                    movel(spat_flatM_pick_p, a=0.2, v=0.1)
                    # begin: URCap Program Node
                    #   Source: Robotiq_Grippers, 3.17.0.105337, Robotiq Inc.
                    #   Type: Gripper
                    $ 4563 "Gripper Open (1)" "noBreak"
                    if not(gripper_connected[0]):
                      popup("Gripper 1 must be connected to run this program.", "No connection", False, True, True)
                    end
                    if not(rq_is_gripper_activated("1")):
                      popup("Gripper 1 is not activated. Go to Installation tab > Gripper to activate it and run the program again.", "Not activated", False, True, True)
                    end
                    rq_set_pos_spd_for(0, 0, 77, "1")
                    rq_wait_pos_spe_for_request(0, 0, 77, "1")
                    rq_go_to("1")
                    rq_wait("1")
                    # end: URCap Program Node
                    $ 4564 "spat_flatS_pick" "noBreak"
                    movel(spat_flatS_pick_p, a=1.2, v=0.25)
                    # begin: URCap Program Node
                    #   Source: Robotiq_Grippers, 3.17.0.105337, Robotiq Inc.
                    #   Type: Gripper
                    $ 4565 "Gripper Close (1)" "noBreak"
                    if not(gripper_connected[0]):
                      popup("Gripper 1 must be connected to run this program.", "No connection", False, True, True)
                    end
                    if not(rq_is_gripper_activated("1")):
                      popup("Gripper 1 is not activated. Go to Installation tab > Gripper to activate it and run the program again.", "Not activated", False, True, True)
                    end
                    rq_set_pos_spd_for(255, 0, 77, "1")
                    rq_wait_pos_spe_for_request(255, 0, 77, "1")
                    rq_go_to("1")
                    rq_wait("1")
                    # end: URCap Program Node
                    $ 4566 "spat_flatS_up" "noBreak"
                    movel(spat_flatS_up_p, a=1.2, v=0.25)
                    $ 4567 "Spatula_otw" "noBreak"
                    movel(Spatula_otw_p, a=1.2, v=0.25)
                    $ 4568 "switch_spat_F_S≔ False " "noBreak"
                    global switch_spat_F_S=  False
                    $ 4569 "correction_reset()" "noBreak"
                    correction_reset()
                  end
                end
              end
            end
            $ 4570 "tilt(level)" "noBreak"
            tilt(level)
            $ 4571 "Action_Info≔'Scooping'" "noBreak"
            global Action_Info="Scooping"
            $ 4572 "auto_tilt_and_scoop(W_now, target_weight, weight_value)" "noBreak"
            auto_tilt_and_scoop(W_now, target_weight, weight_value)
            $ 4573 "Action_Info≔'Dosing'" "noBreak"
            global Action_Info="Dosing"
          end
        end
        if (weight_value <= target_weight and delta_count<3):
          global thread_handler_4490=run Thread_while_4490()
          while (weight_value <= target_weight and delta_count<3):
            sync()
          end
          kill thread_handler_4490
        end
        # begin: URCap Program Node
        #   Source: SensoPart VISOR Robotic, 2.0.6, SensoPart Industriesensorik GmbH
        #   Type: Exit Pose
        $ 4574 "Exit Pose" "noBreak"
        movel(pose_trans(easyPickPose,p[0.0000,0.0000,-0.0000,0.0000,0.0000,0.0000]),a=0.5000,v=0.2500,t=0.000000,r=0.000000)
        # end: URCap Program Node
        easyPickObjTaken = True
      end
      # end: URCap Program Node
      # begin: URCap Program Node
      #   Source: SensoPart VISOR Robotic, 2.0.6, SensoPart Industriesensorik GmbH
      #   Type: No Object Detected
      $ 4575 "No Object Detected" "noBreak"
      if (visor_partsFound(easyPickVisorId) < 1):
        $ 4576 "Popup: No weigh scale detected" "noBreak"
        popup("No weigh scale detected", "Message", False, False, blocking=True)
        else:
      end
      # end: URCap Program Node
    end
    easyPickCount_4 = easyPickCount_4 + 1
    visor_easyPickUpdate(easyPickVisorId, "counter", easyPickCount_4)
    visor_easyPickSetIdent("bfde9f", easyPickVisorId)
    # end: URCap Program Node
  end
  visorFuncEasyPick_8737ac()
  # end: URCap Program Node
  $ 4577 "MoveL"
  $ 4578 "dispense_pos" "breakAfter"
  movel(dispense_pos, a=0.2, v=0.1)
  $ 4580 "Place spatula back to the rack"
  $ 4581 "If spatula ≟ 'spatula_L'"
  if (spatula  ==  "spatula_L"):
    $ 4582 "MoveJ"
    $ 4583 "Spatula_otw" "breakAfter"
    movej(get_inverse_kin(Spatula_otw_p, qnear=Spatula_otw_q), a=1.3962634015954636, v=1.0471975511965976)
    $ 4584 "MoveL"
    $ 4585 "spat_L_up" "breakAfter"
    movel(spat_L_up_p, a=1.2, v=0.25, r=0.05)
    $ 4586 "spat_L_side" "breakAfter"
    movel(spat_L_side_p, a=1.2, v=0.25, r=0.01)
    $ 4587 "spat_L_lift" "breakAfter"
    movel(spat_L_lift_p, a=1.2, v=0.25, r=0.01)
    $ 4588 "spat_L_pick" "breakAfter"
    movel(spat_L_pick_p, a=0.2, v=0.1)
    # begin: URCap Program Node
    #   Source: Robotiq_Grippers, 3.17.0.105337, Robotiq Inc.
    #   Type: Gripper
    $ 4589 "Gripper Open (1)"
    if not(gripper_connected[0]):
      popup("Gripper 1 must be connected to run this program.", "No connection", False, True, True)
    end
    if not(rq_is_gripper_activated("1")):
      popup("Gripper 1 is not activated. Go to Installation tab > Gripper to activate it and run the program again.", "Not activated", False, True, True)
    end
    rq_set_pos_spd_for(0, 128, 128, "1")
    rq_wait_pos_spe_for_request(0, 128, 128, "1")
    rq_go_to("1")
    rq_wait("1")
    # end: URCap Program Node
    $ 4590 "MoveJ"
    $ 4591 "pick_spat_L_abv" "breakAfter"
    movej(get_inverse_kin(pick_spat_L_abv_p, qnear=pick_spat_L_abv_q), a=1.3962634015954636, v=1.0471975511965976)
    $ 4592 "Spatula_otw" "breakAfter"
    movej(get_inverse_kin(Spatula_otw_p, qnear=Spatula_otw_q), a=1.3962634015954636, v=1.0471975511965976)
  else:
    $ 4593 "ElseIf spatula ≟'spatula_M'"
    if (spatula  == "spatula_M"):
      $ 4594 "MoveJ"
      $ 4595 "Spatula_otw" "breakAfter"
      movej(get_inverse_kin(Spatula_otw_p, qnear=Spatula_otw_q), a=1.3962634015954636, v=1.0471975511965976)
      $ 4596 "spat_M_up" "breakAfter"
      movej(get_inverse_kin(spat_M_up_p, qnear=spat_M_up_q), a=1.3962634015954636, v=1.0471975511965976, r=0.05)
      $ 4597 "MoveL"
      $ 4598 "spat_M_pick" "breakAfter"
      movel(spat_M_pick_p, a=0.2, v=0.1)
      # begin: URCap Program Node
      #   Source: Robotiq_Grippers, 3.17.0.105337, Robotiq Inc.
      #   Type: Gripper
      $ 4599 "Gripper Open (1)"
      if not(gripper_connected[0]):
        popup("Gripper 1 must be connected to run this program.", "No connection", False, True, True)
      end
      if not(rq_is_gripper_activated("1")):
        popup("Gripper 1 is not activated. Go to Installation tab > Gripper to activate it and run the program again.", "Not activated", False, True, True)
      end
      rq_set_pos_spd_for(0, 128, 128, "1")
      rq_wait_pos_spe_for_request(0, 128, 128, "1")
      rq_go_to("1")
      rq_wait("1")
      # end: URCap Program Node
      $ 4600 "spat_M_up" "breakAfter"
      movel(spat_M_up_p, a=1.2, v=0.25, r=0.05)
      $ 4601 "Spatula_otw" "breakAfter"
      movel(Spatula_otw_p, a=1.2, v=0.25)
      $ 4602 "switch_spat_M≔ False "
      global switch_spat_M=  False
    else:
      $ 4603 "ElseIf spatula≟'spatula_S'"
      if (spatula == "spatula_S"):
        $ 4604 "MoveJ"
        $ 4605 "Spatula_otw" "breakAfter"
        movej(get_inverse_kin(Spatula_otw_p, qnear=Spatula_otw_q), a=1.3962634015954636, v=1.0471975511965976)
        $ 4606 "spat_S_Up_7" "breakAfter"
        movej(get_inverse_kin(spat_S_Up_7_p, qnear=spat_S_Up_7_q), a=1.3962634015954636, v=1.0471975511965976, r=0.05)
        $ 4607 "MoveL"
        $ 4608 "spat_S_Pick_4" "breakAfter"
        movel(spat_S_Pick_4_p, a=0.2, v=0.1)
        # begin: URCap Program Node
        #   Source: Robotiq_Grippers, 3.17.0.105337, Robotiq Inc.
        #   Type: Gripper
        $ 4609 "Gripper Open (1)"
        if not(gripper_connected[0]):
          popup("Gripper 1 must be connected to run this program.", "No connection", False, True, True)
        end
        if not(rq_is_gripper_activated("1")):
          popup("Gripper 1 is not activated. Go to Installation tab > Gripper to activate it and run the program again.", "Not activated", False, True, True)
        end
        rq_set_pos_spd_for(0, 255, 51, "1")
        rq_wait_pos_spe_for_request(0, 255, 51, "1")
        rq_go_to("1")
        rq_wait("1")
        # end: URCap Program Node
        $ 4610 "spat_S_Up_8" "breakAfter"
        movel(spat_S_Up_8_p, a=1.2, v=0.25, r=0.05)
        $ 4611 "Spatula_otw" "breakAfter"
        movel(Spatula_otw_p, a=1.2, v=0.25)
        $ 4612 "switch_spat_S≔ False "
        global switch_spat_S=  False
      else:
        $ 4613 "ElseIf spatula≟'spatula_flat_M'"
        if (spatula == "spatula_flat_M"):
          $ 4614 "MoveJ"
          $ 4615 "Spatula_otw" "breakAfter"
          movej(get_inverse_kin(Spatula_otw_p, qnear=Spatula_otw_q), a=1.3962634015954636, v=1.0471975511965976)
          $ 4616 "spat_flatM_up" "breakAfter"
          movej(get_inverse_kin(spat_flatM_up_p, qnear=spat_flatM_up_q), a=1.3962634015954636, v=1.0471975511965976, r=0.05)
          $ 4617 "MoveL"
          $ 4618 "spat_flatM_pick" "breakAfter"
          movel(spat_flatM_pick_p, a=0.2, v=0.1)
          # begin: URCap Program Node
          #   Source: Robotiq_Grippers, 3.17.0.105337, Robotiq Inc.
          #   Type: Gripper
          $ 4619 "Gripper Open (1)"
          if not(gripper_connected[0]):
            popup("Gripper 1 must be connected to run this program.", "No connection", False, True, True)
          end
          if not(rq_is_gripper_activated("1")):
            popup("Gripper 1 is not activated. Go to Installation tab > Gripper to activate it and run the program again.", "Not activated", False, True, True)
          end
          rq_set_pos_spd_for(0, 128, 128, "1")
          rq_wait_pos_spe_for_request(0, 128, 128, "1")
          rq_go_to("1")
          rq_wait("1")
          # end: URCap Program Node
          $ 4620 "spat_flatM_up" "breakAfter"
          movel(spat_flatM_up_p, a=1.2, v=0.25, r=0.05)
          $ 4621 "Spatula_otw" "breakAfter"
          movel(Spatula_otw_p, a=1.2, v=0.25)
          $ 4622 "switch_spat_F_M≔ False "
          global switch_spat_F_M=  False
        else:
          $ 4623 "ElseIf spatula≟'spatula_flat_S'"
          if (spatula == "spatula_flat_S"):
            $ 4624 "MoveJ"
            $ 4625 "Spatula_otw" "breakAfter"
            movej(get_inverse_kin(Spatula_otw_p, qnear=Spatula_otw_q), a=1.3962634015954636, v=1.0471975511965976)
            $ 4626 "spat_flatS_up" "breakAfter"
            movej(get_inverse_kin(spat_flatS_up_p, qnear=spat_flatS_up_q), a=1.3962634015954636, v=1.0471975511965976, r=0.05)
            $ 4627 "MoveL"
            $ 4628 "spat_flatS_pick" "breakAfter"
            movel(spat_flatS_pick_p, a=0.2, v=0.1)
            # begin: URCap Program Node
            #   Source: Robotiq_Grippers, 3.17.0.105337, Robotiq Inc.
            #   Type: Gripper
            $ 4629 "Gripper Open (1)"
            if not(gripper_connected[0]):
              popup("Gripper 1 must be connected to run this program.", "No connection", False, True, True)
            end
            if not(rq_is_gripper_activated("1")):
              popup("Gripper 1 is not activated. Go to Installation tab > Gripper to activate it and run the program again.", "Not activated", False, True, True)
            end
            rq_set_pos_spd_for(0, 128, 128, "1")
            rq_wait_pos_spe_for_request(0, 128, 128, "1")
            rq_go_to("1")
            rq_wait("1")
            # end: URCap Program Node
            $ 4630 "spat_flatS_up" "breakAfter"
            movel(spat_flatS_up_p, a=1.2, v=0.25, r=0.05)
            $ 4631 "Spatula_otw" "breakAfter"
            movel(Spatula_otw_p, a=1.2, v=0.25)
            $ 4632 "switch_spat_F_S≔ False "
            global switch_spat_F_S=  False
          end
        end
      end
    end
  end
  $ 4633 "switch_spat_M≔ True "
  global switch_spat_M=  True
  $ 4634 "switch_spat_S≔ True "
  global switch_spat_S=  True
  $ 4635 "switch_spat_F_M≔ True "
  global switch_spat_F_M=  True
  $ 4636 "switch_spat_F_S≔ True "
  global switch_spat_F_S=  True
  elif (51 == switch_1):
    $ 4646 "Case 51"
    $ 4647 "Task≔'Decapping'"
    global Task="Decapping"
    $ 4648 "tilt_to_home()"
    tilt_to_home()
    $ 4649 "Weigh, Place & decap container"
    $ 4650 "Set"
    set_tcp(p[0.0,0.0,0.15052000000000001,3.1415,0.0,0.0])
    # begin: URCap Program Node
    #   Source: SensoPart VISOR Robotic, 2.0.6, SensoPart Industriesensorik GmbH
    #   Type: VISOR Robotic App
    $ 4651 "VISOR Easy Pick"
    def visorFuncEasyPick_00d6e6():
      # begin: URCap Program Node
      #   Source: SensoPart VISOR Robotic, 2.0.6, SensoPart Industriesensorik GmbH
      #   Type: Easy Pick Setup
      $ 4652 "# 1 Setup" "noBreak"
      local easyPickVisorId = 1
      local easyPickArmMounted = True
      local easyPickSetJob = True
      local easyPickJobName = "PoTS"
      local easyPickAtImgAcq = False
      local easyPickImgAcqPose = FRM_PoTS
      # end: URCap Program Node
      # begin: URCap Program Node
      #   Source: SensoPart VISOR Robotic, 2.0.6, SensoPart Industriesensorik GmbH
      #   Type: Process
      $ 4653 "Process" "noBreak"
      local easyPickObjTaken = False
      local easyPickTrigger = False
      local easyPickPoseIdx = 0
      local easyPickPose = p[0,0,0,0,0,0]
      def easyPickFuncTrigger(visorId, setJob, jobName, arm):
      if (setJob):
        visor_changeJob(visorId, jobName, 6000)
      end
      if (arm):
        visor_trigger(visorId, 6000, "arm")
      else:
        visor_trigger(visorId, 6000)
      end
      global easyPickParts_7=visor_partsFound(visorId)
      visor_easyPickUpdate(visorId, "parts", visor_partsFound(visorId))
      return visor_getPose3d(visorId, 0)
    end
    while (not easyPickObjTaken):
      easyPickTrigger = (easyPickCount_7 >= visor_partsFound(easyPickVisorId)) or (easyPickCount_7 > 9) or (not visor_easyPickCheckIdent("6ff59d", easyPickVisorId))
      if (easyPickTrigger):
        easyPickCount_7 = 0
      end
      easyPickPoseIdx = easyPickCount_7
      easyPickPose = visor_getPose3d(easyPickVisorId, easyPickPoseIdx)
      visor_easyPickUpdate(easyPickVisorId, "counter", easyPickPoseIdx)
      # begin: URCap Program Node
      #   Source: SensoPart VISOR Robotic, 2.0.6, SensoPart Industriesensorik GmbH
      #   Type: Image Acquisition Pose
      $ 4654 "Image Acquisition Pose" "noBreak"
      if (easyPickTrigger):
        if (not easyPickAtImgAcq):
          movej(pose_trans(easyPickImgAcqPose,p[0.0000,0.0000,-0.0000,0.0000,0.0000,0.0000]),a=1.3963,v=1.0472,t=0.000000,r=0.000000)
          easyPickAtImgAcq = True
        end
        easyPickPose = easyPickFuncTrigger(easyPickVisorId, easyPickSetJob, easyPickJobName, easyPickArmMounted)
      end
      # end: URCap Program Node
      # begin: URCap Program Node
      #   Source: SensoPart VISOR Robotic, 2.0.6, SensoPart Industriesensorik GmbH
      #   Type: Object Detected
      $ 4655 "Object Detected" "noBreak"
      if (visor_partsFound(easyPickVisorId) > 0):
        $ 4656 "Open Gripper" "noBreak"
        # begin: URCap Program Node
        #   Source: Robotiq_Grippers, 3.17.0.105337, Robotiq Inc.
        #   Type: Gripper
        $ 4657 "Gripper Open (1)" "noBreak"
        if not(gripper_connected[0]):
          popup("Gripper 1 must be connected to run this program.", "No connection", False, True, True)
        end
        if not(rq_is_gripper_activated("1")):
          popup("Gripper 1 is not activated. Go to Installation tab > Gripper to activate it and run the program again.", "Not activated", False, True, True)
        end
        rq_set_pos_spd_for(0, 77, 77, "1")
        rq_wait_pos_spe_for_request(0, 77, 77, "1")
        rq_go_to("1")
        rq_wait("1")
        # end: URCap Program Node
        $ 4658 "Set" "noBreak"
        set_tcp(p[0.0,0.0,0.161,3.1415,0.0,0.0])
        $ 4659 "Wait: 0.2" "noBreak"
        sleep(0.2)
        $ 4660 "Place on second weigh scale" "noBreak"
        $ 4661 "MoveJ" "noBreak"
        $ 4662 "Waypoint_1" "noBreak"
        movej(get_inverse_kin(Waypoint_1_p, qnear=Waypoint_1_q), a=1.3962634015954636, v=1.0471975511965976, r=0.1)
        $ 4663 "Waypoint_5" "noBreak"
        movej(get_inverse_kin(Waypoint_5_p, qnear=Waypoint_5_q), a=1.3962634015954636, v=1.0471975511965976)
        $ 4665 "If Picking≟ True " "noBreak"
        if (Picking ==   True  ):
          $ 4666 "Pick from saved pose" "noBreak"
          $ 4667 "MoveL" "noBreak"
          $ 4668 "cont_B_safe" "noBreak"
          movel(cont_B_safe_p, a=0.2, v=0.1)
          $ 4669 "saved_place_pos" "noBreak"
          movel(saved_place_pos, a=1.2, v=0.25)
          # begin: URCap Program Node
          #   Source: Robotiq_Grippers, 3.17.0.105337, Robotiq Inc.
          #   Type: Gripper
          $ 4670 "Gripper Close (1)" "noBreak"
          if not(gripper_connected[0]):
            popup("Gripper 1 must be connected to run this program.", "No connection", False, True, True)
          end
          if not(rq_is_gripper_activated("1")):
            popup("Gripper 1 is not activated. Go to Installation tab > Gripper to activate it and run the program again.", "Not activated", False, True, True)
          end
          rq_set_pos_spd_for(255, 77, 26, "1")
          rq_wait_pos_spe_for_request(255, 77, 26, "1")
          rq_go_to("1")
          rq_wait("1")
          # end: URCap Program Node
          $ 4671 "cont_B_safe" "noBreak"
          movel(cont_B_safe_p, a=1.2, v=0.25)
          $ 4672 "Postions_otw" "noBreak"
          movel(Postions_otw_p, a=1.2, v=0.25)
        else:
          $ 4675 "Else" "noBreak"
          $ 4676 "read_db_data()" "noBreak"
          read_db_data()
          $ 4677 "Pick from B" "noBreak"
          $ 4678 "MoveL" "noBreak"
          $ 4680 "cont_B_safe" "noBreak"
          movel(cont_B_safe_p, a=1.2, v=0.25)
          $ 4681 "cont_B_prepick≔pose_trans(Cont_B_TCP, p[0,0,cent_edge/2,0,0,0])" "noBreak"
          global cont_B_prepick= pose_trans (Cont_B_TCP, p[0,0,cent_edge/2,0,0,0])
          $ 4682 "cont_B_otw" "noBreak"
          movel(cont_B_otw_p, a=1.2, v=0.25)
          $ 4684 "cont_B_pick≔pose_trans(cont_B_prepick, p[0,pick_2_base-d_cc,0,0,0,0])" "noBreak"
          global cont_B_pick= pose_trans (cont_B_prepick, p[0,pick_2_base-d_cc,0,0,0,0])
          $ 4685 "cont_B_pick" "noBreak"
          movel(cont_B_pick, a=0.2, v=0.1)
          # begin: URCap Program Node
          #   Source: Robotiq_Grippers, 3.17.0.105337, Robotiq Inc.
          #   Type: Gripper
          $ 4686 "Gripper Close (1)" "noBreak"
          if not(gripper_connected[0]):
            popup("Gripper 1 must be connected to run this program.", "No connection", False, True, True)
          end
          if not(rq_is_gripper_activated("1")):
            popup("Gripper 1 is not activated. Go to Installation tab > Gripper to activate it and run the program again.", "Not activated", False, True, True)
          end
          rq_set_pos_spd_for(255, 77, 51, "1")
          rq_wait_pos_spe_for_request(255, 77, 51, "1")
          rq_go_to("1")
          rq_wait("1")
          # end: URCap Program Node
          $ 4687 "cont_B_prepick" "noBreak"
          movel(cont_B_prepick, a=1.2, v=0.25, r=0.01)
          $ 4688 "Postions_otw" "noBreak"
          movel(Postions_otw_p, a=1.2, v=0.25)
        end
        $ 4690 "MoveJ" "noBreak"
        $ 4691 "Waypoint_12" "noBreak"
        movej(get_inverse_kin(Waypoint_12_p, qnear=Waypoint_12_q), a=1.3962634015954636, v=1.0471975511965976)
        $ 4692 "Waypoint_18" "noBreak"
        movej(get_inverse_kin(Waypoint_18_p, qnear=Waypoint_18_q), a=0.6981317007977318, v=0.5235987755982988)
        $ 4693 "w_full_thread≔ True " "noBreak"
        global w_full_thread=  True
        $ 4694 "MoveL" "noBreak"
        $ 4695 "Waypoint_19" "noBreak"
        global move_thread_flag_4695=0
        thread move_thread_4695():
          enter_critical
          move_thread_flag_4695 = 1
          movel(Waypoint_19_p, a=0.2, v=0.005)
          move_thread_flag_4695 = 2
          exit_critical
        end
        move_thread_flag_4695 = 0
        move_thread_han_4695 = run move_thread_4695()
        while (True):
          local targetTcpDirection=get_target_tcp_speed()
          local stepsToRetract=tool_contact(direction=targetTcpDirection, force_threshold=1.000000)
          if (stepsToRetract > 0):
            kill move_thread_han_4695
            stopl(6.0)
            local backTrackMovement=get_actual_joint_positions_history(stepsToRetract)
            local contactPose=get_forward_kin(backTrackMovement)
            local posDir=[targetTcpDirection[0],targetTcpDirection[1],targetTcpDirection[2]]
            local retractTo=contactPose
            if (norm(posDir) > 1e-6):
              local normalizedPosDir=normalize(posDir)
              local additionalRetraction=p[normalizedPosDir[0] * 0.0, normalizedPosDir[1] * 0.0, normalizedPosDir[2] * 0.0, 0, 0, 0]
              retractTo = pose_sub(contactPose, additionalRetraction)
            end
            movel(retractTo, a=6.0, v=0.1)
            $ 4696 "Until (tool_contact_detection)" "noBreak"
            # begin: URCap Program Node
            #   Source: Robotiq_Grippers, 3.17.0.105337, Robotiq Inc.
            #   Type: Gripper
            $ 4697 "Gripper Open (1)" "noBreak"
            if not(gripper_connected[0]):
              popup("Gripper 1 must be connected to run this program.", "No connection", False, True, True)
            end
            if not(rq_is_gripper_activated("1")):
              popup("Gripper 1 is not activated. Go to Installation tab > Gripper to activate it and run the program again.", "Not activated", False, True, True)
            end
            rq_set_pos_spd_for(0, 77, 0, "1")
            rq_wait_pos_spe_for_request(0, 77, 0, "1")
            rq_go_to("1")
            rq_wait("1")
            # end: URCap Program Node
            break
          end
          sleep(1.0E-10)
          if (move_thread_flag_4695 > 1):
            join move_thread_han_4695
            break
          end
          sync()
        end
        $ 4699 "aa_weight_cont≔get_cont_weight()" "noBreak"
        global aa_weight_cont=get_cont_weight()
        $ 4700 "w_full_thread≔ False " "noBreak"
        global w_full_thread=  False
        # begin: URCap Program Node
        #   Source: Robotiq_Grippers, 3.17.0.105337, Robotiq Inc.
        #   Type: Gripper
        $ 4701 "Gripper Close (1)" "noBreak"
        if not(gripper_connected[0]):
          popup("Gripper 1 must be connected to run this program.", "No connection", False, True, True)
        end
        if not(rq_is_gripper_activated("1")):
          popup("Gripper 1 is not activated. Go to Installation tab > Gripper to activate it and run the program again.", "Not activated", False, True, True)
        end
        rq_set_pos_spd_for(255, 77, 0, "1")
        rq_wait_pos_spe_for_request(255, 77, 0, "1")
        rq_go_to("1")
        rq_wait("1")
        # end: URCap Program Node
        $ 4702 "global W_now = aa_weight_cont" "noBreak"
        global W_now = aa_weight_cont
        $ 4703 "Waypoint_18" "noBreak"
        movej(get_inverse_kin(Waypoint_18_p, qnear=Waypoint_18_q), a=1.3962634015954636, v=1.0471975511965976)
        $ 4704 "Waypoint_12" "noBreak"
        movej(get_inverse_kin(Waypoint_12_p, qnear=Waypoint_12_q), a=1.3962634015954636, v=1.0471975511965976)
        $ 4705 "Set" "noBreak"
        set_tcp(p[0.0,0.0,0.15052000000000001,3.1415,0.0,0.0])
        # begin: URCap Program Node
        #   Source: SensoPart VISOR Robotic, 2.0.6, SensoPart Industriesensorik GmbH
        #   Type: Approach Pose
        $ 4706 "Approach Pose" "noBreak"
        movej(pose_trans(easyPickPose,p[0.0000,0.0000,-0.0000,0.0000,0.0000,0.0000]),a=0.5236,v=0.4363,t=0.000000,r=0.000000)
        # end: URCap Program Node
        # begin: URCap Program Node
        #   Source: SensoPart VISOR Robotic, 2.0.6, SensoPart Industriesensorik GmbH
        #   Type: Target Pose
        $ 4707 "Target Pose" "noBreak"
        movel(pose_trans(easyPickPose,p[0.0000,0.0000,-0.0000,0.0000,0.0000,0.0000]),a=0.1000,v=0.0500,t=0.000000,r=0.000000)
        # end: URCap Program Node
        $ 4708 "Close Gripper" "noBreak"
        $ 4709 "container_place≔get_actual_tcp_pose()" "noBreak"
        global container_place= get_actual_tcp_pose ()
        $ 4710 "PoTS_place_abov≔pose_trans(container_place, p[0,0,cent_edge/2,0,0,0])" "noBreak"
        global PoTS_place_abov=pose_trans(container_place, p[0,0,cent_edge/2,0,0,0])
        $ 4711 "MoveL" "noBreak"
        $ 4712 "PoTS_place_abov" "noBreak"
        movel(PoTS_place_abov, a=0.5, v=0.05)
        $ 4714 "target_pose≔pose_trans(PoTS_place_abov, p[0,pick_2_base-d_cc,0,0,0,0])" "noBreak"
        global target_pose=pose_trans(PoTS_place_abov, p[0,pick_2_base-d_cc,0,0,0,0])
        $ 4715 "MoveL" "noBreak"
        $ 4716 "target_pose" "noBreak"
        movel(target_pose, a=0.3, v=0.05)
        # begin: URCap Program Node
        #   Source: Robotiq_Grippers, 3.17.0.105337, Robotiq Inc.
        #   Type: Gripper
        $ 4717 "Gripper Open (1)" "noBreak"
        if not(gripper_connected[0]):
          popup("Gripper 1 must be connected to run this program.", "No connection", False, True, True)
        end
        if not(rq_is_gripper_activated("1")):
          popup("Gripper 1 is not activated. Go to Installation tab > Gripper to activate it and run the program again.", "Not activated", False, True, True)
        end
        rq_set_pos_spd_for(0, 77, 77, "1")
        rq_wait_pos_spe_for_request(0, 77, 77, "1")
        rq_go_to("1")
        rq_wait("1")
        # end: URCap Program Node
        # begin: URCap Program Node
        #   Source: SensoPart VISOR Robotic, 2.0.6, SensoPart Industriesensorik GmbH
        #   Type: Exit Pose
        $ 4718 "Exit Pose" "noBreak"
        movel(pose_trans(easyPickPose,p[0.0000,0.0000,0.1000,0.0000,0.0000,0.0000]),a=0.5000,v=0.2500,t=0.000000,r=0.000000)
        # end: URCap Program Node
        easyPickObjTaken = True
      end
      # end: URCap Program Node
      # begin: URCap Program Node
      #   Source: SensoPart VISOR Robotic, 2.0.6, SensoPart Industriesensorik GmbH
      #   Type: No Object Detected
      $ 4719 "No Object Detected" "noBreak"
      if (visor_partsFound(easyPickVisorId) < 1):
        $ 4720 "Popup: No POTS detected" "noBreak"
        popup("No POTS detected", "Message", False, False, blocking=True)
        else:
      end
      # end: URCap Program Node
    end
    easyPickCount_7 = easyPickCount_7 + 1
    visor_easyPickUpdate(easyPickVisorId, "counter", easyPickCount_7)
    visor_easyPickSetIdent("6ff59d", easyPickVisorId)
    # end: URCap Program Node
  end
  visorFuncEasyPick_00d6e6()
  # end: URCap Program Node
  $ 4721 "Decapping pose"
  $ 4722 "cont_cent_pots=center_pose()"
  cont_cent_pots=center_pose()
  $ 4723 "pre_safe_decap≔pose_trans(cont_cent_pots,p[0,0,0.06,0,0,0])"
  global pre_safe_decap=pose_trans(cont_cent_pots,p[0,0,0.06,0,0,0])
  $ 4724 "decap_pots≔pose_trans(cont_cent_pots,p[0,0,H_c-H+0.02,0,0,0])"
  global decap_pots=pose_trans(cont_cent_pots,p[0,0,H_c-H+0.02,0,0,0])
  $ 4725 "MoveL"
  $ 4726 "MoveJ"
  $ 4727 "FRM_PoTS" "breakAfter"
  movej(FRM_PoTS, a=1.3962634015954636, v=1.0471975511965976)
  $ 4728 "pre_safe_decap" "breakAfter"
  movel(pre_safe_decap, a=0.6, v=0.1)
  $ 4731 "decap_pots" "breakAfter"
  movel(decap_pots, a=0.6, v=0.1)
  # begin: URCap Program Node
  #   Source: Robotiq_Grippers, 3.17.0.105337, Robotiq Inc.
  #   Type: Gripper
  $ 4732 "Gripper Close (1)"
  if not(gripper_connected[0]):
    popup("Gripper 1 must be connected to run this program.", "No connection", False, True, True)
  end
  if not(rq_is_gripper_activated("1")):
    popup("Gripper 1 is not activated. Go to Installation tab > Gripper to activate it and run the program again.", "Not activated", False, True, True)
  end
  rq_set_pos_spd_for(255, 127, 127, "1")
  rq_wait_pos_spe_for_request(255, 127, 127, "1")
  rq_go_to("1")
  rq_wait("1")
  # end: URCap Program Node
  $ 4733 "Decapping"
  $ 4734 "CW_full_Rotate()"
  CW_full_Rotate()
  $ 4735 "CW_full_Rotate()"
  CW_full_Rotate()
  $ 4736 "Wait: 5.0"
  sleep(5.0)
  $ 4737 "decapped≔pose_trans(decap_pots,p[0,0,0.03,0,0,0])"
  global decapped= pose_trans (decap_pots,p[0,0,0.03,0,0,0])
  $ 4740 "MoveL"
  $ 4741 "decapped" "breakAfter"
  movel(decapped, a=0.015, v=0.003)
  $ 4743 "tilt_to_home()"
  tilt_to_home()
  $ 4744 "Placing the cap"
  $ 4745 "pre_cap_place≔pose_trans(pre_safe_decap,p[-0.11,0,0,0,0,-1.5708])"
  global pre_cap_place= pose_trans (pre_safe_decap,p[-0.11,0,0,0,0,-1.5708])
  $ 4746 "pre_cap_place" "breakAfter"
  movel(pre_cap_place, a=0.6, v=0.1)
  $ 4747 "place_cap≔pose_trans(pre_cap_place, p[0,0,-H-0.05,0,0,0])"
  global place_cap= pose_trans (pre_cap_place, p[0,0,-H-0.05,0,0,0])
  $ 4748 "place_cap" "breakAfter"
  global move_thread_flag_4748=0
  thread move_thread_4748():
    enter_critical
    move_thread_flag_4748 = 1
    movel(place_cap, a=0.2, v=0.1)
    move_thread_flag_4748 = 2
    exit_critical
  end
  move_thread_flag_4748 = 0
  move_thread_han_4748 = run move_thread_4748()
  while (True):
    local targetTcpDirection=get_target_tcp_speed()
    local stepsToRetract=tool_contact(direction=targetTcpDirection, force_threshold=1.000000)
    if (stepsToRetract > 0):
      kill move_thread_han_4748
      stopl(5.0)
      local backTrackMovement=get_actual_joint_positions_history(stepsToRetract)
      local contactPose=get_forward_kin(backTrackMovement)
      local posDir=[targetTcpDirection[0],targetTcpDirection[1],targetTcpDirection[2]]
      local retractTo=contactPose
      if (norm(posDir) > 1e-6):
        local normalizedPosDir=normalize(posDir)
        local additionalRetraction=p[normalizedPosDir[0] * 1.0E-4, normalizedPosDir[1] * 1.0E-4, normalizedPosDir[2] * 1.0E-4, 0, 0, 0]
        retractTo = pose_sub(contactPose, additionalRetraction)
      end
      movel(retractTo, a=5.0, v=0.1)
      $ 4749 "Until (tool_contact_detection)"
      $ 4750 "Cap_pose≔get_actual_tcp_pose()"
      global Cap_pose= get_actual_tcp_pose ()
      break
    end
    sleep(1.0E-10)
    if (move_thread_flag_4748 > 1):
      join move_thread_han_4748
      break
    end
    sync()
  end
  # begin: URCap Program Node
  #   Source: Robotiq_Grippers, 3.17.0.105337, Robotiq Inc.
  #   Type: Gripper
  $ 4751 "Gripper Open (1)"
  if not(gripper_connected[0]):
    popup("Gripper 1 must be connected to run this program.", "No connection", False, True, True)
  end
  if not(rq_is_gripper_activated("1")):
    popup("Gripper 1 is not activated. Go to Installation tab > Gripper to activate it and run the program again.", "Not activated", False, True, True)
  end
  rq_set_pos_spd_for(0, 255, 77, "1")
  rq_wait_pos_spe_for_request(0, 255, 77, "1")
  rq_go_to("1")
  rq_wait("1")
  # end: URCap Program Node
  $ 4752 "pre_cap_place" "breakAfter"
  movel(pre_cap_place, a=0.6, v=0.1)
  $ 4755 "MoveJ"
  $ 4756 "place_2_home" "breakAfter"
  movej(get_inverse_kin(place_2_home_p, qnear=place_2_home_q), a=1.3962634015954636, v=1.0471975511965976)
  $ 4757 "Picking≔ False "
  global Picking=  False
  elif (52 == switch_1):
    $ 4758 "Case 52"
    $ 4759 "Task≔'Dosing'"
    global Task="Dosing"
    $ 4760 "tilt_to_home()"
    tilt_to_home()
    $ 4761 "Powder dosing all"
    $ 4762 "tilt_angle_sent≔0.0"
    global tilt_angle_sent=0.0
    $ 4763 "send_target_info()"
    send_target_info()
    $ 4765 "prev_spat≔''"
    global prev_spat=""
    $ 4766 "spatula≔''"
    global spatula=""
    $ 4767 "scoop_status≔'normal'"
    global scoop_status="normal"
    $ 4768 "send_powder_info()"
    send_powder_info()
    $ 4769 "Set AO[0]=0.0"
    set_standard_analog_out(0, 0.0)
    $ 4770 "Wait: 0.2"
    sleep(0.2)
    $ 4771 "reach pots decapping pose"
    # begin: URCap Program Node
    #   Source: SensoPart VISOR Robotic, 2.0.6, SensoPart Industriesensorik GmbH
    #   Type: VISOR Robotic App
    $ 4777 "VISOR Easy Pick"
    def visorFuncEasyPick_00f506():
      # begin: URCap Program Node
      #   Source: SensoPart VISOR Robotic, 2.0.6, SensoPart Industriesensorik GmbH
      #   Type: Easy Pick Setup
      $ 4778 "# 1 Setup" "noBreak"
      local easyPickVisorId = 1
      local easyPickArmMounted = True
      local easyPickSetJob = True
      local easyPickJobName = "Weight_scale"
      local easyPickAtImgAcq = False
      local easyPickImgAcqPose = Trigger
      # end: URCap Program Node
      # begin: URCap Program Node
      #   Source: SensoPart VISOR Robotic, 2.0.6, SensoPart Industriesensorik GmbH
      #   Type: Process
      $ 4779 "Process" "noBreak"
      local easyPickObjTaken = False
      local easyPickTrigger = False
      local easyPickPoseIdx = 0
      local easyPickPose = p[0,0,0,0,0,0]
      def easyPickFuncTrigger(visorId, setJob, jobName, arm):
      if (setJob):
        visor_changeJob(visorId, jobName, 6000)
      end
      if (arm):
        visor_trigger(visorId, 6000, "arm")
      else:
        visor_trigger(visorId, 6000)
      end
      global easyPickParts_4=visor_partsFound(visorId)
      visor_easyPickUpdate(visorId, "parts", visor_partsFound(visorId))
      return visor_getPose3d(visorId, 0)
    end
    while (not easyPickObjTaken):
      easyPickTrigger = (easyPickCount_4 >= visor_partsFound(easyPickVisorId)) or (easyPickCount_4 > 9) or (not visor_easyPickCheckIdent("4fb698", easyPickVisorId))
      if (easyPickTrigger):
        easyPickCount_4 = 0
      end
      easyPickPoseIdx = easyPickCount_4
      easyPickPose = visor_getPose3d(easyPickVisorId, easyPickPoseIdx)
      visor_easyPickUpdate(easyPickVisorId, "counter", easyPickPoseIdx)
      # begin: URCap Program Node
      #   Source: SensoPart VISOR Robotic, 2.0.6, SensoPart Industriesensorik GmbH
      #   Type: Image Acquisition Pose
      $ 4780 "Image Acquisition Pose" "noBreak"
      if (easyPickTrigger):
        if (not easyPickAtImgAcq):
          movej(pose_trans(easyPickImgAcqPose,p[0.0000,0.0000,-0.0000,0.0000,0.0000,0.0000]),a=1.3963,v=1.0472,t=0.000000,r=0.000000)
          easyPickAtImgAcq = True
        end
        easyPickPose = easyPickFuncTrigger(easyPickVisorId, easyPickSetJob, easyPickJobName, easyPickArmMounted)
      end
      # end: URCap Program Node
      # begin: URCap Program Node
      #   Source: SensoPart VISOR Robotic, 2.0.6, SensoPart Industriesensorik GmbH
      #   Type: Object Detected
      $ 4781 "Object Detected" "noBreak"
      if (visor_partsFound(easyPickVisorId) > 0):
        $ 4782 "Open Gripper" "noBreak"
        $ 4783 "weight_value≔get_weight()" "noBreak"
        global weight_value=get_weight()
        $ 4784 "Wait: 0.5" "noBreak"
        sleep(0.5)
        $ 4785 "diff≔target_weight-weight_value" "noBreak"
        global diff=target_weight-weight_value
        $ 4786 "compute_level_percent(W_now, weight_value)" "noBreak"
        compute_level_percent(W_now, weight_value)
        $ 4787 "send_level_info()" "noBreak"
        send_level_info()
        $ 4788 "spatula≔select_spatula(Flowability, level, diff, bulk_density, mouth_d)" "noBreak"
        global spatula=select_spatula(Flowability, level, diff, bulk_density, mouth_d)
        $ 4789 "Wait: 0.2" "noBreak"
        sleep(0.2)
        $ 4790 "send_spatula_info()" "noBreak"
        send_spatula_info()
        $ 4791 "Pick spatula" "noBreak"
        $ 4792 "If spatula ≟ 'spatula_L'" "noBreak"
        if (spatula  ==  "spatula_L"):
          $ 4793 "MoveJ" "noBreak"
          $ 4794 "Spatula_otw" "noBreak"
          movej(get_inverse_kin(Spatula_otw_p, qnear=Spatula_otw_q), a=1.3962634015954636, v=1.0471975511965976)
          $ 4795 "pick_spat_L_abv" "noBreak"
          movej(get_inverse_kin(pick_spat_L_abv_p, qnear=pick_spat_L_abv_q), a=1.3962634015954636, v=1.0471975511965976)
          $ 4796 "MoveL" "noBreak"
          $ 4797 "spat_L_pick" "noBreak"
          movel(spat_L_pick_p, a=1.2, v=0.25)
          # begin: URCap Program Node
          #   Source: Robotiq_Grippers, 3.17.0.105337, Robotiq Inc.
          #   Type: Gripper
          $ 4798 "Gripper Close (1)" "noBreak"
          if not(gripper_connected[0]):
            popup("Gripper 1 must be connected to run this program.", "No connection", False, True, True)
          end
          if not(rq_is_gripper_activated("1")):
            popup("Gripper 1 is not activated. Go to Installation tab > Gripper to activate it and run the program again.", "Not activated", False, True, True)
          end
          rq_set_pos_spd_for(255, 0, 77, "1")
          rq_wait_pos_spe_for_request(255, 0, 77, "1")
          rq_go_to("1")
          rq_wait("1")
          # end: URCap Program Node
          $ 4799 "spat_L_lift" "noBreak"
          movel(spat_L_lift_p, a=1.2, v=0.25, r=0.01)
          $ 4800 "spat_L_side" "noBreak"
          movel(spat_L_side_p, a=1.2, v=0.25, r=0.01)
          $ 4801 "spat_L_up" "noBreak"
          movel(spat_L_up_p, a=1.2, v=0.25, r=0.05)
          $ 4802 "MoveJ" "noBreak"
          $ 4803 "Spatula_otw" "noBreak"
          movej(get_inverse_kin(Spatula_otw_p, qnear=Spatula_otw_q), a=1.3962634015954636, v=1.0471975511965976)
        else:
          $ 4804 "ElseIf spatula ≟'spatula_M'" "noBreak"
          if (spatula  == "spatula_M"):
            $ 4805 "MoveJ" "noBreak"
            $ 4806 "Spatula_otw" "noBreak"
            movej(get_inverse_kin(Spatula_otw_p, qnear=Spatula_otw_q), a=1.3962634015954636, v=1.0471975511965976)
            $ 4807 "spat_M_up" "noBreak"
            movej(get_inverse_kin(spat_M_up_p, qnear=spat_M_up_q), a=1.3962634015954636, v=1.0471975511965976, r=0.05)
            $ 4808 "MoveL" "noBreak"
            $ 4809 "spat_M_pick" "noBreak"
            movel(spat_M_pick_p, a=1.2, v=0.25)
            # begin: URCap Program Node
            #   Source: Robotiq_Grippers, 3.17.0.105337, Robotiq Inc.
            #   Type: Gripper
            $ 4810 "Gripper Close (1)" "noBreak"
            if not(gripper_connected[0]):
              popup("Gripper 1 must be connected to run this program.", "No connection", False, True, True)
            end
            if not(rq_is_gripper_activated("1")):
              popup("Gripper 1 is not activated. Go to Installation tab > Gripper to activate it and run the program again.", "Not activated", False, True, True)
            end
            rq_set_pos_spd_for(255, 0, 77, "1")
            rq_wait_pos_spe_for_request(255, 0, 77, "1")
            rq_go_to("1")
            rq_wait("1")
            # end: URCap Program Node
            $ 4811 "spat_M_up" "noBreak"
            movel(spat_M_up_p, a=1.2, v=0.25, r=0.05)
            $ 4812 "Spatula_otw" "noBreak"
            movel(Spatula_otw_p, a=1.2, v=0.25)
            $ 4813 "switch_spat_M≔ False " "noBreak"
            global switch_spat_M=  False
          else:
            $ 4814 "ElseIf spatula≟'spatula_S'" "noBreak"
            if (spatula == "spatula_S"):
              $ 4815 "MoveJ" "noBreak"
              $ 4816 "Spatula_otw" "noBreak"
              movej(get_inverse_kin(Spatula_otw_p, qnear=Spatula_otw_q), a=1.3962634015954636, v=1.0471975511965976)
              $ 4817 "spat_S_Up_7" "noBreak"
              movej(get_inverse_kin(spat_S_Up_7_p, qnear=spat_S_Up_7_q), a=1.3962634015954636, v=1.0471975511965976, r=0.05)
              $ 4818 "MoveL" "noBreak"
              $ 4819 "spat_S_Pick_4" "noBreak"
              movel(spat_S_Pick_4_p, a=1.2, v=0.25)
              # begin: URCap Program Node
              #   Source: Robotiq_Grippers, 3.17.0.105337, Robotiq Inc.
              #   Type: Gripper
              $ 4820 "Gripper Close (1)" "noBreak"
              if not(gripper_connected[0]):
                popup("Gripper 1 must be connected to run this program.", "No connection", False, True, True)
              end
              if not(rq_is_gripper_activated("1")):
                popup("Gripper 1 is not activated. Go to Installation tab > Gripper to activate it and run the program again.", "Not activated", False, True, True)
              end
              rq_set_pos_spd_for(255, 0, 77, "1")
              rq_wait_pos_spe_for_request(255, 0, 77, "1")
              rq_go_to("1")
              rq_wait("1")
              # end: URCap Program Node
              $ 4821 "spat_S_Up_8" "noBreak"
              movel(spat_S_Up_8_p, a=1.2, v=0.25, r=0.05)
              $ 4822 "Spatula_otw" "noBreak"
              movel(Spatula_otw_p, a=1.2, v=0.25)
              $ 4823 "switch_spat_S≔ False " "noBreak"
              global switch_spat_S=  False
            else:
              $ 4824 "ElseIf spatula≟'spatula_flat_M'" "noBreak"
              if (spatula == "spatula_flat_M"):
                $ 4825 "MoveJ" "noBreak"
                $ 4826 "Spatula_otw" "noBreak"
                movej(get_inverse_kin(Spatula_otw_p, qnear=Spatula_otw_q), a=1.3962634015954636, v=1.0471975511965976)
                $ 4827 "spat_flatM_up" "noBreak"
                movej(get_inverse_kin(spat_flatM_up_p, qnear=spat_flatM_up_q), a=1.3962634015954636, v=1.0471975511965976, r=0.05)
                $ 4828 "MoveL" "noBreak"
                $ 4829 "spat_flatM_pick" "noBreak"
                movel(spat_flatM_pick_p, a=1.2, v=0.25)
                # begin: URCap Program Node
                #   Source: Robotiq_Grippers, 3.17.0.105337, Robotiq Inc.
                #   Type: Gripper
                $ 4830 "Gripper Close (1)" "noBreak"
                if not(gripper_connected[0]):
                  popup("Gripper 1 must be connected to run this program.", "No connection", False, True, True)
                end
                if not(rq_is_gripper_activated("1")):
                  popup("Gripper 1 is not activated. Go to Installation tab > Gripper to activate it and run the program again.", "Not activated", False, True, True)
                end
                rq_set_pos_spd_for(255, 0, 77, "1")
                rq_wait_pos_spe_for_request(255, 0, 77, "1")
                rq_go_to("1")
                rq_wait("1")
                # end: URCap Program Node
                $ 4831 "spat_flatM_up" "noBreak"
                movel(spat_flatM_up_p, a=1.2, v=0.25, r=0.05)
                $ 4832 "Spatula_otw" "noBreak"
                movel(Spatula_otw_p, a=1.2, v=0.25)
                $ 4833 "switch_spat_F_M≔ False " "noBreak"
                global switch_spat_F_M=  False
              else:
                $ 4834 "ElseIf spatula≟'spatula_flat_S'" "noBreak"
                if (spatula == "spatula_flat_S"):
                  $ 4835 "MoveJ" "noBreak"
                  $ 4836 "Spatula_otw" "noBreak"
                  movej(get_inverse_kin(Spatula_otw_p, qnear=Spatula_otw_q), a=1.3962634015954636, v=1.0471975511965976)
                  $ 4837 "spat_flatS_up" "noBreak"
                  movej(get_inverse_kin(spat_flatS_up_p, qnear=spat_flatS_up_q), a=1.3962634015954636, v=1.0471975511965976, r=0.05)
                  $ 4838 "MoveL" "noBreak"
                  $ 4839 "spat_flatS_pick" "noBreak"
                  movel(spat_flatS_pick_p, a=1.2, v=0.25)
                  # begin: URCap Program Node
                  #   Source: Robotiq_Grippers, 3.17.0.105337, Robotiq Inc.
                  #   Type: Gripper
                  $ 4840 "Gripper Close (1)" "noBreak"
                  if not(gripper_connected[0]):
                    popup("Gripper 1 must be connected to run this program.", "No connection", False, True, True)
                  end
                  if not(rq_is_gripper_activated("1")):
                    popup("Gripper 1 is not activated. Go to Installation tab > Gripper to activate it and run the program again.", "Not activated", False, True, True)
                  end
                  rq_set_pos_spd_for(255, 0, 77, "1")
                  rq_wait_pos_spe_for_request(255, 0, 77, "1")
                  rq_go_to("1")
                  rq_wait("1")
                  # end: URCap Program Node
                  $ 4841 "spat_flatS_up" "noBreak"
                  movel(spat_flatS_up_p, a=1.2, v=0.25, r=0.05)
                  $ 4842 "Spatula_otw" "noBreak"
                  movel(Spatula_otw_p, a=1.2, v=0.25)
                  $ 4843 "switch_spat_F_S≔ False " "noBreak"
                  global switch_spat_F_S=  False
                end
              end
            end
          end
        end
        $ 4844 "Action_Info≔'Scooping'" "noBreak"
        global Action_Info="Scooping"
        $ 4845 "auto_tilt_and_scoop(W_now, target_weight, weight_value)" "noBreak"
        auto_tilt_and_scoop(W_now, target_weight, weight_value)
        $ 4846 "Action_Info≔'Dosing'" "noBreak"
        global Action_Info="Dosing"
        # begin: URCap Program Node
        #   Source: SensoPart VISOR Robotic, 2.0.6, SensoPart Industriesensorik GmbH
        #   Type: Approach Pose
        $ 4847 "Approach Pose" "noBreak"
        movej(pose_trans(easyPickPose,p[0.0000,0.0000,-0.0000,0.0000,0.0000,0.0000]),a=0.2618,v=0.1745,t=0.000000,r=0.000000)
        # end: URCap Program Node
        # begin: URCap Program Node
        #   Source: SensoPart VISOR Robotic, 2.0.6, SensoPart Industriesensorik GmbH
        #   Type: Target Pose
        $ 4848 "Target Pose" "noBreak"
        movel(pose_trans(easyPickPose,p[0.0000,0.0000,-0.0000,0.0000,0.0000,0.0000]),a=0.0500,v=0.0200,t=0.000000,r=0.000000)
        # end: URCap Program Node
        $ 4849 "Close Gripper" "noBreak"
        $ 4850 "current_p≔get_actual_tcp_pose()" "noBreak"
        global current_p= get_actual_tcp_pose ()
        $ 4851 "dispense_pos≔pose_trans(current_p,p[0,0,0,0,-deg2rad(spatula_ry),0])" "noBreak"
        global dispense_pos=pose_trans(current_p,p[0,0,0,0,-deg2rad(spatula_ry),0])
        $ 4852 "Loop weight_value≤target_weight and delta_count≤3" "noBreak"
        thread Thread_while_4852():
          while (True):
            $ 4853 "MoveL" "noBreak"
            $ 4854 "dispense_pos" "noBreak"
            movel(dispense_pos, a=0.2, v=0.1)
            $ 4855 "log_weight()" "noBreak"
            log_weight()
            $ 4857 "CCW_full_Rotate()" "noBreak"
            CCW_full_Rotate()
            $ 4858 "Start_thread≔ True " "noBreak"
            global Start_thread=  True
            $ 4859 "vib_thread≔ True " "noBreak"
            global vib_thread=  True
            $ 4860 "Wait: 0.5" "noBreak"
            sleep(0.5)
            $ 4861 "If diff ≥(target_g*1.2)" "noBreak"
            if (diff  >= (target_g*1.2)):
              $ 4862 "tilt_pose≔pose_trans(get_actual_tcp_pose(), p[0, 0, 0, 0, 0, 2.0])" "noBreak"
              global tilt_pose=pose_trans(get_actual_tcp_pose(), p[0, 0, 0, 0, 0, 2.0])
              $ 4863 "movel(tilt_pose, a=0.5, v=0.5, r=0.00001)" "noBreak"
              movel(tilt_pose, a=0.5, v=0.5, r=0.00001)
            else:
              $ 4864 "Else" "noBreak"
              $ 4865 "Loop weight_value≤(target_weight-0.00) and tilt_angle≥(-1.999) and tilt_angle≤0.5" "noBreak"
              thread Thread_while_4865():
                while (True):
                  $ 4866 "current_error≔target_weight-weight_value" "noBreak"
                  global current_error=target_weight-weight_value
                  $ 4867 "Integral_error≔Integral_error+current_error*dt" "noBreak"
                  global Integral_error=Integral_error+current_error*dt
                  $ 4868 "derivative≔(current_error-previous_error)/dt" "noBreak"
                  global derivative=(current_error-previous_error)/dt
                  $ 4869 "tilt_increment≔(kp*current_error)+(ki*Integral_error)+(kd*derivative)" "noBreak"
                  global tilt_increment=(kp*current_error)+(ki*Integral_error)+(kd*derivative)
                  $ 4870 "current_pose≔get_actual_tcp_pose()" "noBreak"
                  global current_pose= get_actual_tcp_pose ()
                  $ 4871 "tilt_angle≔current_pose[5]" "noBreak"
                  global tilt_angle=current_pose[5]
                  $ 4872 "tilt_pose≔pose_trans(current_pose, p[0, 0, 0, 0, 0, tilt_increment])" "noBreak"
                  global tilt_pose=pose_trans(current_pose, p[0, 0, 0, 0, 0, tilt_increment])
                  $ 4873 "movel(tilt_pose, a=0.1, v=0.1, r=0.00001)" "noBreak"
                  movel(tilt_pose, a=0.1, v=0.1, r=0.00001)
                  $ 4874 "previous_error≔current_error" "noBreak"
                  global previous_error=current_error
                end
              end
              if (weight_value <= (target_weight-0.00)  and  tilt_angle >= (-1.999)  and  tilt_angle <= 0.5):
                global thread_handler_4865=run Thread_while_4865()
                while (weight_value <= (target_weight-0.00)  and  tilt_angle >= (-1.999)  and  tilt_angle <= 0.5):
                  sync()
                end
                kill thread_handler_4865
              end
            end
            $ 4875 "weight_value≔get_weight()" "noBreak"
            global weight_value=get_weight()
            $ 4876 "tilt_angle≔-1" "noBreak"
            global tilt_angle=-1
            $ 4877 "Wait: 0.5" "noBreak"
            sleep(0.5)
            $ 4878 "Start_thread≔ False " "noBreak"
            global Start_thread=  False
            $ 4879 "vib_thread≔ False " "noBreak"
            global vib_thread=  False
            $ 4880 "dispense_pos" "noBreak"
            movel(dispense_pos, a=1.2, v=0.25)
            $ 4881 "compute_level_percent(W_now, weight_value)" "noBreak"
            compute_level_percent(W_now, weight_value)
            $ 4882 "If delta<0.01" "noBreak"
            if (delta<0.01):
              $ 4883 "delta_count≔delta_count+1" "noBreak"
              global delta_count=delta_count+1
            else:
              $ 4884 "Else" "noBreak"
              $ 4885 "delta_count≔0" "noBreak"
              global delta_count=0
            end
            $ 4886 "prev_spat≔spatula" "noBreak"
            global prev_spat=spatula
            $ 4887 "Wait: 0.2" "noBreak"
            sleep(0.2)
            $ 4888 "spatula≔select_spatula(Flowability, level, diff, bulk_density, mouth_d)" "noBreak"
            global spatula=select_spatula(Flowability, level, diff, bulk_density, mouth_d)
            $ 4889 "Wait: 1.0" "noBreak"
            sleep(1.0)
            $ 4890 "send_level_info()" "noBreak"
            send_level_info()
            $ 4891 "send_spatula_info()" "noBreak"
            send_spatula_info()
            $ 4892 "Integral_error≔0" "noBreak"
            global Integral_error=0
            $ 4893 "current_error≔0" "noBreak"
            global current_error=0
            $ 4894 "previous_error≔0" "noBreak"
            global previous_error=0
            $ 4895 "Set AO[0]=0.0" "noBreak"
            set_standard_analog_out(0, 0.0)
            $ 4896 "Wait: 0.5" "noBreak"
            sleep(0.5)
            $ 4897 "swtich spatula" "noBreak"
            $ 4898 "If spatula ≟ 'spatula_M' and switch_spat_M≟ True " "noBreak"
            if (spatula  ==  "spatula_M"  and  switch_spat_M ==   True  ):
              $ 4899 "MoveJ" "noBreak"
              $ 4900 "Spatula_otw" "noBreak"
              movej(get_inverse_kin(Spatula_otw_p, qnear=Spatula_otw_q), a=1.3962634015954636, v=1.0471975511965976)
              $ 4901 "spat_L_up" "noBreak"
              movej(get_inverse_kin(spat_L_up_p, qnear=spat_L_up_q), a=1.3962634015954636, v=1.0471975511965976)
              $ 4902 "MoveL" "noBreak"
              $ 4903 "spat_L_side" "noBreak"
              movel(spat_L_side_p, a=1.2, v=0.25)
              $ 4904 "spat_L_lift" "noBreak"
              movel(spat_L_lift_p, a=1.2, v=0.25)
              $ 4905 "spat_L_pick" "noBreak"
              movel(spat_L_pick_p, a=0.2, v=0.1)
              # begin: URCap Program Node
              #   Source: Robotiq_Grippers, 3.17.0.105337, Robotiq Inc.
              #   Type: Gripper
              $ 4906 "Gripper Open (1)" "noBreak"
              if not(gripper_connected[0]):
                popup("Gripper 1 must be connected to run this program.", "No connection", False, True, True)
              end
              if not(rq_is_gripper_activated("1")):
                popup("Gripper 1 is not activated. Go to Installation tab > Gripper to activate it and run the program again.", "Not activated", False, True, True)
              end
              rq_set_pos_spd_for(0, 255, 77, "1")
              rq_wait_pos_spe_for_request(0, 255, 77, "1")
              rq_go_to("1")
              rq_wait("1")
              # end: URCap Program Node
              $ 4907 "spat_M_pick" "noBreak"
              movel(spat_M_pick_p, a=1.2, v=0.25)
              # begin: URCap Program Node
              #   Source: Robotiq_Grippers, 3.17.0.105337, Robotiq Inc.
              #   Type: Gripper
              $ 4908 "Gripper Close (1)" "noBreak"
              if not(gripper_connected[0]):
                popup("Gripper 1 must be connected to run this program.", "No connection", False, True, True)
              end
              if not(rq_is_gripper_activated("1")):
                popup("Gripper 1 is not activated. Go to Installation tab > Gripper to activate it and run the program again.", "Not activated", False, True, True)
              end
              rq_set_pos_spd_for(255, 0, 77, "1")
              rq_wait_pos_spe_for_request(255, 0, 77, "1")
              rq_go_to("1")
              rq_wait("1")
              # end: URCap Program Node
              $ 4909 "spat_M_up" "noBreak"
              movel(spat_M_up_p, a=1.2, v=0.25)
              $ 4910 "Spatula_otw" "noBreak"
              movel(Spatula_otw_p, a=1.2, v=0.25)
              $ 4911 "switch_spat_M≔ False " "noBreak"
              global switch_spat_M=  False
              $ 4912 "correction_reset()" "noBreak"
              correction_reset()
            else:
              $ 4913 "ElseIf spatula ≟ 'spatula_S' and switch_spat_S ≟ True and prev_spat≟'spatula_M'" "noBreak"
              if (spatula  ==  "spatula_S" and switch_spat_S  ==   True  and prev_spat == "spatula_M"):
                $ 4914 "MoveL" "noBreak"
                $ 4915 "Spatula_otw" "noBreak"
                movel(Spatula_otw_p, a=1.2, v=0.25)
                $ 4916 "spat_M_up" "noBreak"
                movel(spat_M_up_p, a=1.2, v=0.25)
                $ 4917 "spat_M_pick" "noBreak"
                movel(spat_M_pick_p, a=0.2, v=0.1)
                # begin: URCap Program Node
                #   Source: Robotiq_Grippers, 3.17.0.105337, Robotiq Inc.
                #   Type: Gripper
                $ 4918 "Gripper Open (1)" "noBreak"
                if not(gripper_connected[0]):
                  popup("Gripper 1 must be connected to run this program.", "No connection", False, True, True)
                end
                if not(rq_is_gripper_activated("1")):
                  popup("Gripper 1 is not activated. Go to Installation tab > Gripper to activate it and run the program again.", "Not activated", False, True, True)
                end
                rq_set_pos_spd_for(0, 255, 77, "1")
                rq_wait_pos_spe_for_request(0, 255, 77, "1")
                rq_go_to("1")
                rq_wait("1")
                # end: URCap Program Node
                $ 4919 "spat_S_pick" "noBreak"
                movel(spat_S_pick_p, a=1.2, v=0.25)
                # begin: URCap Program Node
                #   Source: Robotiq_Grippers, 3.17.0.105337, Robotiq Inc.
                #   Type: Gripper
                $ 4920 "Gripper Close (1)" "noBreak"
                if not(gripper_connected[0]):
                  popup("Gripper 1 must be connected to run this program.", "No connection", False, True, True)
                end
                if not(rq_is_gripper_activated("1")):
                  popup("Gripper 1 is not activated. Go to Installation tab > Gripper to activate it and run the program again.", "Not activated", False, True, True)
                end
                rq_set_pos_spd_for(255, 0, 77, "1")
                rq_wait_pos_spe_for_request(255, 0, 77, "1")
                rq_go_to("1")
                rq_wait("1")
                # end: URCap Program Node
                $ 4921 "spat_S_up" "noBreak"
                movel(spat_S_up_p, a=1.2, v=0.25)
                $ 4922 "Spatula_otw" "noBreak"
                movel(Spatula_otw_p, a=1.2, v=0.25)
                $ 4923 "switch_spat_S≔ False " "noBreak"
                global switch_spat_S=  False
                $ 4924 "correction_reset()" "noBreak"
                correction_reset()
              else:
                $ 4925 "ElseIf spatula≟'spatula_S' and switch_spat_S≟ True  and prev_spat≟'spatula_L'" "noBreak"
                if (spatula == "spatula_S" and switch_spat_S ==   True    and  prev_spat == "spatula_L"):
                  $ 4926 "MoveJ" "noBreak"
                  $ 4927 "Spatula_otw" "noBreak"
                  movej(get_inverse_kin(Spatula_otw_p, qnear=Spatula_otw_q), a=1.3962634015954636, v=1.0471975511965976)
                  $ 4928 "spat_L_up" "noBreak"
                  movej(get_inverse_kin(spat_L_up_p, qnear=spat_L_up_q), a=1.3962634015954636, v=1.0471975511965976)
                  $ 4929 "MoveL" "noBreak"
                  $ 4930 "spat_L_side" "noBreak"
                  movel(spat_L_side_p, a=1.2, v=0.25)
                  $ 4931 "spat_L_lift" "noBreak"
                  movel(spat_L_lift_p, a=1.2, v=0.25)
                  $ 4932 "spat_L_pick" "noBreak"
                  movel(spat_L_pick_p, a=0.2, v=0.1)
                  # begin: URCap Program Node
                  #   Source: Robotiq_Grippers, 3.17.0.105337, Robotiq Inc.
                  #   Type: Gripper
                  $ 4933 "Gripper Open (1)" "noBreak"
                  if not(gripper_connected[0]):
                    popup("Gripper 1 must be connected to run this program.", "No connection", False, True, True)
                  end
                  if not(rq_is_gripper_activated("1")):
                    popup("Gripper 1 is not activated. Go to Installation tab > Gripper to activate it and run the program again.", "Not activated", False, True, True)
                  end
                  rq_set_pos_spd_for(0, 255, 77, "1")
                  rq_wait_pos_spe_for_request(0, 255, 77, "1")
                  rq_go_to("1")
                  rq_wait("1")
                  # end: URCap Program Node
                  $ 4934 "spat_S_pick" "noBreak"
                  movel(spat_S_pick_p, a=1.2, v=0.25)
                  # begin: URCap Program Node
                  #   Source: Robotiq_Grippers, 3.17.0.105337, Robotiq Inc.
                  #   Type: Gripper
                  $ 4935 "Gripper Close (1)" "noBreak"
                  if not(gripper_connected[0]):
                    popup("Gripper 1 must be connected to run this program.", "No connection", False, True, True)
                  end
                  if not(rq_is_gripper_activated("1")):
                    popup("Gripper 1 is not activated. Go to Installation tab > Gripper to activate it and run the program again.", "Not activated", False, True, True)
                  end
                  rq_set_pos_spd_for(255, 0, 77, "1")
                  rq_wait_pos_spe_for_request(255, 0, 77, "1")
                  rq_go_to("1")
                  rq_wait("1")
                  # end: URCap Program Node
                  $ 4936 "spat_S_up" "noBreak"
                  movel(spat_S_up_p, a=1.2, v=0.25)
                  $ 4937 "Spatula_otw" "noBreak"
                  movel(Spatula_otw_p, a=1.2, v=0.25)
                  $ 4938 "switch_spat_S≔ False " "noBreak"
                  global switch_spat_S=  False
                  $ 4939 "correction_reset()" "noBreak"
                  correction_reset()
                else:
                  $ 4940 "ElseIf spatula≟'spatula_flat_S'  and switch_spat_F_S ≟ True " "noBreak"
                  if (spatula == "spatula_flat_S"   and  switch_spat_F_S  ==   True  ):
                    $ 4941 "MoveL" "noBreak"
                    $ 4942 "Spatula_otw" "noBreak"
                    movel(Spatula_otw_p, a=1.2, v=0.25)
                    $ 4943 "spat_flatM_up" "noBreak"
                    movel(spat_flatM_up_p, a=1.2, v=0.25)
                    $ 4944 "spat_flatM_pick" "noBreak"
                    movel(spat_flatM_pick_p, a=0.2, v=0.1)
                    # begin: URCap Program Node
                    #   Source: Robotiq_Grippers, 3.17.0.105337, Robotiq Inc.
                    #   Type: Gripper
                    $ 4945 "Gripper Open (1)" "noBreak"
                    if not(gripper_connected[0]):
                      popup("Gripper 1 must be connected to run this program.", "No connection", False, True, True)
                    end
                    if not(rq_is_gripper_activated("1")):
                      popup("Gripper 1 is not activated. Go to Installation tab > Gripper to activate it and run the program again.", "Not activated", False, True, True)
                    end
                    rq_set_pos_spd_for(0, 255, 74, "1")
                    rq_wait_pos_spe_for_request(0, 255, 74, "1")
                    rq_go_to("1")
                    rq_wait("1")
                    # end: URCap Program Node
                    $ 4946 "spat_flatS_pick" "noBreak"
                    movel(spat_flatS_pick_p, a=1.2, v=0.25)
                    # begin: URCap Program Node
                    #   Source: Robotiq_Grippers, 3.17.0.105337, Robotiq Inc.
                    #   Type: Gripper
                    $ 4947 "Gripper Close (1)" "noBreak"
                    if not(gripper_connected[0]):
                      popup("Gripper 1 must be connected to run this program.", "No connection", False, True, True)
                    end
                    if not(rq_is_gripper_activated("1")):
                      popup("Gripper 1 is not activated. Go to Installation tab > Gripper to activate it and run the program again.", "Not activated", False, True, True)
                    end
                    rq_set_pos_spd_for(255, 0, 77, "1")
                    rq_wait_pos_spe_for_request(255, 0, 77, "1")
                    rq_go_to("1")
                    rq_wait("1")
                    # end: URCap Program Node
                    $ 4948 "spat_flatS_up" "noBreak"
                    movel(spat_flatS_up_p, a=1.2, v=0.25)
                    $ 4949 "Spatula_otw" "noBreak"
                    movel(Spatula_otw_p, a=1.2, v=0.25)
                    $ 4950 "switch_spat_F_S≔ False " "noBreak"
                    global switch_spat_F_S=  False
                    $ 4951 "correction_reset()" "noBreak"
                    correction_reset()
                  end
                end
              end
            end
            $ 4952 "tilt(level)" "noBreak"
            tilt(level)
            $ 4953 "Action_Info≔'Scooping'" "noBreak"
            global Action_Info="Scooping"
            $ 4954 "auto_tilt_and_scoop(W_now, target_weight, weight_value)" "noBreak"
            auto_tilt_and_scoop(W_now, target_weight, weight_value)
            $ 4955 "Action_Info≔'Dosing'" "noBreak"
            global Action_Info="Dosing"
          end
        end
        if (weight_value <= target_weight and delta_count <= 3):
          global thread_handler_4852=run Thread_while_4852()
          while (weight_value <= target_weight and delta_count <= 3):
            sync()
          end
          kill thread_handler_4852
        end
        $ 4956 "Start_thread≔ False " "noBreak"
        global Start_thread=  False
        $ 4957 "vib_thread≔ False " "noBreak"
        global vib_thread=  False
        # begin: URCap Program Node
        #   Source: SensoPart VISOR Robotic, 2.0.6, SensoPart Industriesensorik GmbH
        #   Type: Exit Pose
        $ 4958 "Exit Pose" "noBreak"
        movel(pose_trans(easyPickPose,p[0.0000,0.0000,-0.0000,0.0000,0.0000,0.0000]),a=0.5000,v=0.2500,t=0.000000,r=0.000000)
        # end: URCap Program Node
        easyPickObjTaken = True
      end
      # end: URCap Program Node
      # begin: URCap Program Node
      #   Source: SensoPart VISOR Robotic, 2.0.6, SensoPart Industriesensorik GmbH
      #   Type: No Object Detected
      $ 4959 "No Object Detected" "noBreak"
      if (visor_partsFound(easyPickVisorId) < 1):
        $ 4960 "Popup: No weigh scale detected" "noBreak"
        popup("No weigh scale detected", "Message", False, False, blocking=True)
        else:
      end
      # end: URCap Program Node
    end
    easyPickCount_4 = easyPickCount_4 + 1
    visor_easyPickUpdate(easyPickVisorId, "counter", easyPickCount_4)
    visor_easyPickSetIdent("4fb698", easyPickVisorId)
    # end: URCap Program Node
  end
  visorFuncEasyPick_00f506()
  # end: URCap Program Node
  $ 4961 "MoveL"
  $ 4962 "dispense_pos" "breakAfter"
  movel(dispense_pos, a=0.2, v=0.1)
  $ 4963 "after_scoop()"
  after_scoop()
  $ 4964 "Place spatula back to the rack"
  $ 4965 "If spatula ≟ 'spatula_L'"
  if (spatula  ==  "spatula_L"):
    $ 4966 "MoveJ"
    $ 4967 "Spatula_otw" "breakAfter"
    movej(get_inverse_kin(Spatula_otw_p, qnear=Spatula_otw_q), a=1.3962634015954636, v=1.0471975511965976)
    $ 4968 "MoveL"
    $ 4969 "spat_L_up" "breakAfter"
    movel(spat_L_up_p, a=1.2, v=0.25, r=0.05)
    $ 4970 "spat_L_side" "breakAfter"
    movel(spat_L_side_p, a=1.2, v=0.25, r=0.01)
    $ 4971 "spat_L_lift" "breakAfter"
    movel(spat_L_lift_p, a=1.2, v=0.25, r=0.01)
    $ 4972 "spat_L_pick" "breakAfter"
    movel(spat_L_pick_p, a=0.2, v=0.1)
    # begin: URCap Program Node
    #   Source: Robotiq_Grippers, 3.17.0.105337, Robotiq Inc.
    #   Type: Gripper
    $ 4973 "Gripper Open (1)"
    if not(gripper_connected[0]):
      popup("Gripper 1 must be connected to run this program.", "No connection", False, True, True)
    end
    if not(rq_is_gripper_activated("1")):
      popup("Gripper 1 is not activated. Go to Installation tab > Gripper to activate it and run the program again.", "Not activated", False, True, True)
    end
    rq_set_pos_spd_for(0, 128, 128, "1")
    rq_wait_pos_spe_for_request(0, 128, 128, "1")
    rq_go_to("1")
    rq_wait("1")
    # end: URCap Program Node
    $ 4974 "MoveJ"
    $ 4975 "pick_spat_L_abv" "breakAfter"
    movej(get_inverse_kin(pick_spat_L_abv_p, qnear=pick_spat_L_abv_q), a=1.3962634015954636, v=1.0471975511965976)
    $ 4976 "Spatula_otw" "breakAfter"
    movej(get_inverse_kin(Spatula_otw_p, qnear=Spatula_otw_q), a=1.3962634015954636, v=1.0471975511965976)
  else:
    $ 4977 "ElseIf spatula ≟'spatula_M'"
    if (spatula  == "spatula_M"):
      $ 4978 "MoveJ"
      $ 4979 "Spatula_otw" "breakAfter"
      movej(get_inverse_kin(Spatula_otw_p, qnear=Spatula_otw_q), a=1.3962634015954636, v=1.0471975511965976)
      $ 4980 "spat_M_up" "breakAfter"
      movej(get_inverse_kin(spat_M_up_p, qnear=spat_M_up_q), a=1.3962634015954636, v=1.0471975511965976, r=0.05)
      $ 4981 "MoveL"
      $ 4982 "spat_M_pick" "breakAfter"
      movel(spat_M_pick_p, a=0.2, v=0.1)
      # begin: URCap Program Node
      #   Source: Robotiq_Grippers, 3.17.0.105337, Robotiq Inc.
      #   Type: Gripper
      $ 4983 "Gripper Open (1)"
      if not(gripper_connected[0]):
        popup("Gripper 1 must be connected to run this program.", "No connection", False, True, True)
      end
      if not(rq_is_gripper_activated("1")):
        popup("Gripper 1 is not activated. Go to Installation tab > Gripper to activate it and run the program again.", "Not activated", False, True, True)
      end
      rq_set_pos_spd_for(0, 128, 128, "1")
      rq_wait_pos_spe_for_request(0, 128, 128, "1")
      rq_go_to("1")
      rq_wait("1")
      # end: URCap Program Node
      $ 4984 "spat_M_up" "breakAfter"
      movel(spat_M_up_p, a=1.2, v=0.25, r=0.05)
      $ 4985 "Spatula_otw" "breakAfter"
      movel(Spatula_otw_p, a=1.2, v=0.25)
      $ 4986 "switch_spat_M≔ False "
      global switch_spat_M=  False
    else:
      $ 4987 "ElseIf spatula≟'spatula_S'"
      if (spatula == "spatula_S"):
        $ 4988 "MoveJ"
        $ 4989 "Spatula_otw" "breakAfter"
        movej(get_inverse_kin(Spatula_otw_p, qnear=Spatula_otw_q), a=1.3962634015954636, v=1.0471975511965976)
        $ 4990 "spat_S_Up_7" "breakAfter"
        movej(get_inverse_kin(spat_S_Up_7_p, qnear=spat_S_Up_7_q), a=1.3962634015954636, v=1.0471975511965976, r=0.05)
        $ 4991 "MoveL"
        $ 4992 "spat_S_Pick_4" "breakAfter"
        movel(spat_S_Pick_4_p, a=0.2, v=0.1)
        # begin: URCap Program Node
        #   Source: Robotiq_Grippers, 3.17.0.105337, Robotiq Inc.
        #   Type: Gripper
        $ 4993 "Gripper Open (1)"
        if not(gripper_connected[0]):
          popup("Gripper 1 must be connected to run this program.", "No connection", False, True, True)
        end
        if not(rq_is_gripper_activated("1")):
          popup("Gripper 1 is not activated. Go to Installation tab > Gripper to activate it and run the program again.", "Not activated", False, True, True)
        end
        rq_set_pos_spd_for(0, 255, 51, "1")
        rq_wait_pos_spe_for_request(0, 255, 51, "1")
        rq_go_to("1")
        rq_wait("1")
        # end: URCap Program Node
        $ 4994 "spat_S_Up_8" "breakAfter"
        movel(spat_S_Up_8_p, a=1.2, v=0.25, r=0.05)
        $ 4995 "Spatula_otw" "breakAfter"
        movel(Spatula_otw_p, a=1.2, v=0.25)
        $ 4996 "switch_spat_S≔ False "
        global switch_spat_S=  False
      else:
        $ 4997 "ElseIf spatula≟'spatula_flat_M'"
        if (spatula == "spatula_flat_M"):
          $ 4998 "MoveJ"
          $ 4999 "Spatula_otw" "breakAfter"
          movej(get_inverse_kin(Spatula_otw_p, qnear=Spatula_otw_q), a=1.3962634015954636, v=1.0471975511965976)
          $ 5000 "spat_flatM_up" "breakAfter"
          movej(get_inverse_kin(spat_flatM_up_p, qnear=spat_flatM_up_q), a=1.3962634015954636, v=1.0471975511965976, r=0.05)
          $ 5001 "MoveL"
          $ 5002 "spat_flatM_pick" "breakAfter"
          movel(spat_flatM_pick_p, a=0.2, v=0.1)
          # begin: URCap Program Node
          #   Source: Robotiq_Grippers, 3.17.0.105337, Robotiq Inc.
          #   Type: Gripper
          $ 5003 "Gripper Open (1)"
          if not(gripper_connected[0]):
            popup("Gripper 1 must be connected to run this program.", "No connection", False, True, True)
          end
          if not(rq_is_gripper_activated("1")):
            popup("Gripper 1 is not activated. Go to Installation tab > Gripper to activate it and run the program again.", "Not activated", False, True, True)
          end
          rq_set_pos_spd_for(0, 128, 128, "1")
          rq_wait_pos_spe_for_request(0, 128, 128, "1")
          rq_go_to("1")
          rq_wait("1")
          # end: URCap Program Node
          $ 5004 "spat_flatM_up" "breakAfter"
          movel(spat_flatM_up_p, a=1.2, v=0.25, r=0.05)
          $ 5005 "Spatula_otw" "breakAfter"
          movel(Spatula_otw_p, a=1.2, v=0.25)
          $ 5006 "switch_spat_F_M≔ False "
          global switch_spat_F_M=  False
        else:
          $ 5007 "ElseIf spatula≟'spatula_flat_S'"
          if (spatula == "spatula_flat_S"):
            $ 5008 "MoveJ"
            $ 5009 "Spatula_otw" "breakAfter"
            movej(get_inverse_kin(Spatula_otw_p, qnear=Spatula_otw_q), a=1.3962634015954636, v=1.0471975511965976)
            $ 5010 "spat_flatS_up" "breakAfter"
            movej(get_inverse_kin(spat_flatS_up_p, qnear=spat_flatS_up_q), a=1.3962634015954636, v=1.0471975511965976, r=0.05)
            $ 5011 "MoveL"
            $ 5012 "spat_flatS_pick" "breakAfter"
            movel(spat_flatS_pick_p, a=0.2, v=0.1)
            # begin: URCap Program Node
            #   Source: Robotiq_Grippers, 3.17.0.105337, Robotiq Inc.
            #   Type: Gripper
            $ 5013 "Gripper Open (1)"
            if not(gripper_connected[0]):
              popup("Gripper 1 must be connected to run this program.", "No connection", False, True, True)
            end
            if not(rq_is_gripper_activated("1")):
              popup("Gripper 1 is not activated. Go to Installation tab > Gripper to activate it and run the program again.", "Not activated", False, True, True)
            end
            rq_set_pos_spd_for(0, 128, 128, "1")
            rq_wait_pos_spe_for_request(0, 128, 128, "1")
            rq_go_to("1")
            rq_wait("1")
            # end: URCap Program Node
            $ 5014 "spat_flatS_up" "breakAfter"
            movel(spat_flatS_up_p, a=1.2, v=0.25, r=0.05)
            $ 5015 "Spatula_otw" "breakAfter"
            movel(Spatula_otw_p, a=1.2, v=0.25)
            $ 5016 "switch_spat_F_S≔ False "
            global switch_spat_F_S=  False
          end
        end
      end
    end
  end
  $ 5017 "switch_spat_M≔ True "
  global switch_spat_M=  True
  $ 5018 "switch_spat_S≔ True "
  global switch_spat_S=  True
  $ 5019 "switch_spat_F_M≔ True "
  global switch_spat_F_M=  True
  $ 5020 "switch_spat_F_S≔ True "
  global switch_spat_F_S=  True
  $ 5021 "correction_reset()"
  correction_reset()
  elif (54 == switch_1):
    $ 5031 "Case 54"
    $ 5032 "Task≔'Fumehood_dosing'"
    global Task="Fumehood_dosing"
    $ 5033 "Powder dosing fumehood"
    $ 5034 "Set"
    set_tcp(p[0.0,0.0,0.15052000000000001,3.1415,0.0,0.0])
    $ 5035 "prev_spat≔''"
    global prev_spat=""
    $ 5036 "spatula≔''"
    global spatula=""
    $ 5037 "scoop_status≔'normal'"
    global scoop_status="normal"
    $ 5038 "Set AO[0]=0.0"
    set_standard_analog_out(0, 0.0)
    $ 5039 "Wait: 0.2"
    sleep(0.2)
    # begin: URCap Program Node
    #   Source: SensoPart VISOR Robotic, 2.0.6, SensoPart Industriesensorik GmbH
    #   Type: VISOR Robotic App
    $ 5040 "VISOR Easy Pick"
    def visorFuncEasyPick_dd8337():
      # begin: URCap Program Node
      #   Source: SensoPart VISOR Robotic, 2.0.6, SensoPart Industriesensorik GmbH
      #   Type: Easy Pick Setup
      $ 5041 "# 1 Setup" "noBreak"
      local easyPickVisorId = 1
      local easyPickArmMounted = True
      local easyPickSetJob = True
      local easyPickJobName = "Fumehood_container"
      local easyPickAtImgAcq = False
      local easyPickImgAcqPose = FRM_PoTS
      # end: URCap Program Node
      # begin: URCap Program Node
      #   Source: SensoPart VISOR Robotic, 2.0.6, SensoPart Industriesensorik GmbH
      #   Type: Process
      $ 5042 "Process" "noBreak"
      local easyPickObjTaken = False
      local easyPickTrigger = False
      local easyPickPoseIdx = 0
      local easyPickPose = p[0,0,0,0,0,0]
      def easyPickFuncTrigger(visorId, setJob, jobName, arm):
      if (setJob):
        visor_changeJob(visorId, jobName, 6000)
      end
      if (arm):
        visor_trigger(visorId, 6000, "arm")
      else:
        visor_trigger(visorId, 6000)
      end
      global easyPickParts_4=visor_partsFound(visorId)
      visor_easyPickUpdate(visorId, "parts", visor_partsFound(visorId))
      return visor_getPose3d(visorId, 0)
    end
    while (not easyPickObjTaken):
      easyPickTrigger = (easyPickCount_4 >= visor_partsFound(easyPickVisorId)) or (easyPickCount_4 > 9) or (not visor_easyPickCheckIdent("3af2be", easyPickVisorId))
      if (easyPickTrigger):
        easyPickCount_4 = 0
      end
      easyPickPoseIdx = easyPickCount_4
      easyPickPose = visor_getPose3d(easyPickVisorId, easyPickPoseIdx)
      visor_easyPickUpdate(easyPickVisorId, "counter", easyPickPoseIdx)
      # begin: URCap Program Node
      #   Source: SensoPart VISOR Robotic, 2.0.6, SensoPart Industriesensorik GmbH
      #   Type: Image Acquisition Pose
      $ 5043 "Image Acquisition Pose" "noBreak"
      if (easyPickTrigger):
        if (not easyPickAtImgAcq):
          movej(pose_trans(easyPickImgAcqPose,p[0.0000,0.0000,-0.0000,0.0000,0.0000,0.0000]),a=1.3963,v=1.0472,t=0.000000,r=0.000000)
          easyPickAtImgAcq = True
        end
        easyPickPose = easyPickFuncTrigger(easyPickVisorId, easyPickSetJob, easyPickJobName, easyPickArmMounted)
      end
      # end: URCap Program Node
      # begin: URCap Program Node
      #   Source: SensoPart VISOR Robotic, 2.0.6, SensoPart Industriesensorik GmbH
      #   Type: Object Detected
      $ 5044 "Object Detected" "noBreak"
      if (visor_partsFound(easyPickVisorId) > 0):
        $ 5045 "Open Gripper" "noBreak"
        $ 5046 "MoveJ" "noBreak"
        $ 5047 "Scan_db" "noBreak"
        movej(get_inverse_kin(Scan_db_p, qnear=Scan_db_q), a=1.3962634015954636, v=1.0471975511965976)
        $ 5048 "read_db_data()" "noBreak"
        read_db_data()
        $ 5049 "read_spatula_data()" "noBreak"
        read_spatula_data()
        $ 5050 "spatula≔'spatula_M'" "noBreak"
        global spatula="spatula_M"
        $ 5051 "Pick spatula" "noBreak"
        $ 5052 "Set" "noBreak"
        set_tcp(p[0.0,0.0,0.161,3.1415,0.0,0.0])
        $ 5053 "If spatula ≟ 'spatula_L'" "noBreak"
        if (spatula  ==  "spatula_L"):
          $ 5054 "MoveJ" "noBreak"
          $ 5055 "Spatula_otw" "noBreak"
          movej(get_inverse_kin(Spatula_otw_p, qnear=Spatula_otw_q), a=1.3962634015954636, v=1.0471975511965976)
          $ 5056 "pick_spat_L_abv" "noBreak"
          movej(get_inverse_kin(pick_spat_L_abv_p, qnear=pick_spat_L_abv_q), a=1.3962634015954636, v=1.0471975511965976)
          $ 5057 "MoveL" "noBreak"
          $ 5058 "spat_L_pick" "noBreak"
          movel(spat_L_pick_p, a=1.2, v=0.25)
          # begin: URCap Program Node
          #   Source: Robotiq_Grippers, 3.17.0.105337, Robotiq Inc.
          #   Type: Gripper
          $ 5059 "Gripper Close (1)" "noBreak"
          if not(gripper_connected[0]):
            popup("Gripper 1 must be connected to run this program.", "No connection", False, True, True)
          end
          if not(rq_is_gripper_activated("1")):
            popup("Gripper 1 is not activated. Go to Installation tab > Gripper to activate it and run the program again.", "Not activated", False, True, True)
          end
          rq_set_pos_spd_for(255, 0, 77, "1")
          rq_wait_pos_spe_for_request(255, 0, 77, "1")
          rq_go_to("1")
          rq_wait("1")
          # end: URCap Program Node
          $ 5060 "spat_L_lift" "noBreak"
          movel(spat_L_lift_p, a=1.2, v=0.25, r=0.01)
          $ 5061 "spat_L_side" "noBreak"
          movel(spat_L_side_p, a=1.2, v=0.25, r=0.01)
          $ 5062 "spat_L_up" "noBreak"
          movel(spat_L_up_p, a=1.2, v=0.25, r=0.05)
          $ 5063 "MoveJ" "noBreak"
          $ 5064 "Spatula_otw" "noBreak"
          movej(get_inverse_kin(Spatula_otw_p, qnear=Spatula_otw_q), a=1.3962634015954636, v=1.0471975511965976)
        else:
          $ 5065 "ElseIf spatula ≟'spatula_M'" "noBreak"
          if (spatula  == "spatula_M"):
            $ 5066 "MoveJ" "noBreak"
            $ 5067 "Spatula_otw" "noBreak"
            movej(get_inverse_kin(Spatula_otw_p, qnear=Spatula_otw_q), a=1.3962634015954636, v=1.0471975511965976)
            $ 5068 "spat_M_up" "noBreak"
            movej(get_inverse_kin(spat_M_up_p, qnear=spat_M_up_q), a=1.3962634015954636, v=1.0471975511965976, r=0.05)
            $ 5069 "MoveL" "noBreak"
            $ 5070 "spat_M_pick" "noBreak"
            movel(spat_M_pick_p, a=1.2, v=0.25)
            # begin: URCap Program Node
            #   Source: Robotiq_Grippers, 3.17.0.105337, Robotiq Inc.
            #   Type: Gripper
            $ 5071 "Gripper Close (1)" "noBreak"
            if not(gripper_connected[0]):
              popup("Gripper 1 must be connected to run this program.", "No connection", False, True, True)
            end
            if not(rq_is_gripper_activated("1")):
              popup("Gripper 1 is not activated. Go to Installation tab > Gripper to activate it and run the program again.", "Not activated", False, True, True)
            end
            rq_set_pos_spd_for(255, 0, 77, "1")
            rq_wait_pos_spe_for_request(255, 0, 77, "1")
            rq_go_to("1")
            rq_wait("1")
            # end: URCap Program Node
            $ 5072 "spat_M_up" "noBreak"
            movel(spat_M_up_p, a=1.2, v=0.25, r=0.05)
            $ 5073 "Spatula_otw" "noBreak"
            movel(Spatula_otw_p, a=1.2, v=0.25)
            $ 5074 "switch_spat_M≔ False " "noBreak"
            global switch_spat_M=  False
          else:
            $ 5075 "ElseIf spatula≟'spatula_S'" "noBreak"
            if (spatula == "spatula_S"):
              $ 5076 "MoveJ" "noBreak"
              $ 5077 "Spatula_otw" "noBreak"
              movej(get_inverse_kin(Spatula_otw_p, qnear=Spatula_otw_q), a=1.3962634015954636, v=1.0471975511965976)
              $ 5078 "spat_S_Up_7" "noBreak"
              movej(get_inverse_kin(spat_S_Up_7_p, qnear=spat_S_Up_7_q), a=1.3962634015954636, v=1.0471975511965976, r=0.05)
              $ 5079 "MoveL" "noBreak"
              $ 5080 "spat_S_Pick_4" "noBreak"
              movel(spat_S_Pick_4_p, a=1.2, v=0.25)
              # begin: URCap Program Node
              #   Source: Robotiq_Grippers, 3.17.0.105337, Robotiq Inc.
              #   Type: Gripper
              $ 5081 "Gripper Close (1)" "noBreak"
              if not(gripper_connected[0]):
                popup("Gripper 1 must be connected to run this program.", "No connection", False, True, True)
              end
              if not(rq_is_gripper_activated("1")):
                popup("Gripper 1 is not activated. Go to Installation tab > Gripper to activate it and run the program again.", "Not activated", False, True, True)
              end
              rq_set_pos_spd_for(255, 0, 77, "1")
              rq_wait_pos_spe_for_request(255, 0, 77, "1")
              rq_go_to("1")
              rq_wait("1")
              # end: URCap Program Node
              $ 5082 "spat_S_Up_8" "noBreak"
              movel(spat_S_Up_8_p, a=1.2, v=0.25, r=0.05)
              $ 5083 "Spatula_otw" "noBreak"
              movel(Spatula_otw_p, a=1.2, v=0.25)
              $ 5084 "switch_spat_S≔ False " "noBreak"
              global switch_spat_S=  False
            else:
              $ 5085 "ElseIf spatula≟'spatula_flat_M'" "noBreak"
              if (spatula == "spatula_flat_M"):
                $ 5086 "MoveJ" "noBreak"
                $ 5087 "Spatula_otw" "noBreak"
                movej(get_inverse_kin(Spatula_otw_p, qnear=Spatula_otw_q), a=1.3962634015954636, v=1.0471975511965976)
                $ 5088 "spat_flatM_up" "noBreak"
                movej(get_inverse_kin(spat_flatM_up_p, qnear=spat_flatM_up_q), a=1.3962634015954636, v=1.0471975511965976, r=0.05)
                $ 5089 "MoveL" "noBreak"
                $ 5090 "spat_flatM_pick" "noBreak"
                movel(spat_flatM_pick_p, a=1.2, v=0.25)
                # begin: URCap Program Node
                #   Source: Robotiq_Grippers, 3.17.0.105337, Robotiq Inc.
                #   Type: Gripper
                $ 5091 "Gripper Close (1)" "noBreak"
                if not(gripper_connected[0]):
                  popup("Gripper 1 must be connected to run this program.", "No connection", False, True, True)
                end
                if not(rq_is_gripper_activated("1")):
                  popup("Gripper 1 is not activated. Go to Installation tab > Gripper to activate it and run the program again.", "Not activated", False, True, True)
                end
                rq_set_pos_spd_for(255, 0, 77, "1")
                rq_wait_pos_spe_for_request(255, 0, 77, "1")
                rq_go_to("1")
                rq_wait("1")
                # end: URCap Program Node
                $ 5092 "spat_flatM_up" "noBreak"
                movel(spat_flatM_up_p, a=1.2, v=0.25, r=0.05)
                $ 5093 "Spatula_otw" "noBreak"
                movel(Spatula_otw_p, a=1.2, v=0.25)
                $ 5094 "switch_spat_F_M≔ False " "noBreak"
                global switch_spat_F_M=  False
              else:
                $ 5095 "ElseIf spatula≟'spatula_flat_S'" "noBreak"
                if (spatula == "spatula_flat_S"):
                  $ 5096 "MoveJ" "noBreak"
                  $ 5097 "Spatula_otw" "noBreak"
                  movej(get_inverse_kin(Spatula_otw_p, qnear=Spatula_otw_q), a=1.3962634015954636, v=1.0471975511965976)
                  $ 5098 "spat_flatS_up" "noBreak"
                  movej(get_inverse_kin(spat_flatS_up_p, qnear=spat_flatS_up_q), a=1.3962634015954636, v=1.0471975511965976, r=0.05)
                  $ 5099 "MoveL" "noBreak"
                  $ 5100 "spat_flatS_pick" "noBreak"
                  movel(spat_flatS_pick_p, a=1.2, v=0.25)
                  # begin: URCap Program Node
                  #   Source: Robotiq_Grippers, 3.17.0.105337, Robotiq Inc.
                  #   Type: Gripper
                  $ 5101 "Gripper Close (1)" "noBreak"
                  if not(gripper_connected[0]):
                    popup("Gripper 1 must be connected to run this program.", "No connection", False, True, True)
                  end
                  if not(rq_is_gripper_activated("1")):
                    popup("Gripper 1 is not activated. Go to Installation tab > Gripper to activate it and run the program again.", "Not activated", False, True, True)
                  end
                  rq_set_pos_spd_for(255, 0, 77, "1")
                  rq_wait_pos_spe_for_request(255, 0, 77, "1")
                  rq_go_to("1")
                  rq_wait("1")
                  # end: URCap Program Node
                  $ 5102 "spat_flatS_up" "noBreak"
                  movel(spat_flatS_up_p, a=1.2, v=0.25, r=0.05)
                  $ 5103 "Spatula_otw" "noBreak"
                  movel(Spatula_otw_p, a=1.2, v=0.25)
                  $ 5104 "switch_spat_F_S≔ False " "noBreak"
                  global switch_spat_F_S=  False
                end
              end
            end
          end
        end
        $ 5105 "Set" "noBreak"
        set_tcp(p[0.0,0.0,0.15052000000000001,3.1415,0.0,0.0])
        # begin: URCap Program Node
        #   Source: SensoPart VISOR Robotic, 2.0.6, SensoPart Industriesensorik GmbH
        #   Type: Approach Pose
        $ 5106 "Approach Pose" "noBreak"
        movej(pose_trans(easyPickPose,p[0.0000,0.0000,0.0500,0.0000,0.0000,0.0000]),a=1.3963,v=1.0472,t=0.000000,r=0.000000)
        # end: URCap Program Node
        # begin: URCap Program Node
        #   Source: SensoPart VISOR Robotic, 2.0.6, SensoPart Industriesensorik GmbH
        #   Type: Target Pose
        $ 5107 "Target Pose" "noBreak"
        movel(pose_trans(easyPickPose,p[0.0000,0.0000,-0.0000,0.0000,0.0000,0.0000]),a=0.0500,v=0.0200,t=0.000000,r=0.000000)
        # end: URCap Program Node
        $ 5108 "Close Gripper" "noBreak"
        $ 5109 "f_center≔get_actual_tcp_pose()" "noBreak"
        global f_center= get_actual_tcp_pose ()
        $ 5110 "Loop 2 times" "noBreak"
        Loop_28 = 0
        while (Loop_28 < 2):
          $ 5113 "auto_scoop(W_now)" "noBreak"
          auto_scoop(W_now)
          $ 5114 "Wait: 0.5" "noBreak"
          sleep(0.5)
          $ 5115 "Set AO[0]=0.0" "noBreak"
          set_standard_analog_out(0, 0.0)
          Loop_28 = Loop_28 + 1
        end
        $ 5116 "prev_spat≔spatula" "noBreak"
        global prev_spat=spatula
        $ 5117 "Wait: 0.5" "noBreak"
        sleep(0.5)
        $ 5118 "spatula≔'spatula_S'" "noBreak"
        global spatula="spatula_S"
        $ 5119 "swtich spatula" "noBreak"
        $ 5120 "Set" "noBreak"
        set_tcp(p[0.0,0.0,0.161,3.1415,0.0,0.0])
        $ 5121 "If spatula ≟ 'spatula_M' and switch_spat_M≟ True " "noBreak"
        if (spatula  ==  "spatula_M"  and  switch_spat_M ==   True  ):
          $ 5122 "MoveJ" "noBreak"
          $ 5123 "Spatula_otw" "noBreak"
          movej(get_inverse_kin(Spatula_otw_p, qnear=Spatula_otw_q), a=1.3962634015954636, v=1.0471975511965976)
          $ 5124 "spat_L_up" "noBreak"
          movej(get_inverse_kin(spat_L_up_p, qnear=spat_L_up_q), a=1.3962634015954636, v=1.0471975511965976)
          $ 5125 "MoveL" "noBreak"
          $ 5126 "spat_L_side" "noBreak"
          movel(spat_L_side_p, a=1.2, v=0.25)
          $ 5127 "spat_L_lift" "noBreak"
          movel(spat_L_lift_p, a=1.2, v=0.25)
          $ 5128 "spat_L_pick" "noBreak"
          movel(spat_L_pick_p, a=0.2, v=0.1)
          # begin: URCap Program Node
          #   Source: Robotiq_Grippers, 3.17.0.105337, Robotiq Inc.
          #   Type: Gripper
          $ 5129 "Gripper Open (1)" "noBreak"
          if not(gripper_connected[0]):
            popup("Gripper 1 must be connected to run this program.", "No connection", False, True, True)
          end
          if not(rq_is_gripper_activated("1")):
            popup("Gripper 1 is not activated. Go to Installation tab > Gripper to activate it and run the program again.", "Not activated", False, True, True)
          end
          rq_set_pos_spd_for(0, 255, 77, "1")
          rq_wait_pos_spe_for_request(0, 255, 77, "1")
          rq_go_to("1")
          rq_wait("1")
          # end: URCap Program Node
          $ 5130 "spat_M_pick" "noBreak"
          movel(spat_M_pick_p, a=1.2, v=0.25)
          # begin: URCap Program Node
          #   Source: Robotiq_Grippers, 3.17.0.105337, Robotiq Inc.
          #   Type: Gripper
          $ 5131 "Gripper Close (1)" "noBreak"
          if not(gripper_connected[0]):
            popup("Gripper 1 must be connected to run this program.", "No connection", False, True, True)
          end
          if not(rq_is_gripper_activated("1")):
            popup("Gripper 1 is not activated. Go to Installation tab > Gripper to activate it and run the program again.", "Not activated", False, True, True)
          end
          rq_set_pos_spd_for(255, 0, 77, "1")
          rq_wait_pos_spe_for_request(255, 0, 77, "1")
          rq_go_to("1")
          rq_wait("1")
          # end: URCap Program Node
          $ 5132 "spat_M_up" "noBreak"
          movel(spat_M_up_p, a=1.2, v=0.25)
          $ 5133 "Spatula_otw" "noBreak"
          movel(Spatula_otw_p, a=1.2, v=0.25)
          $ 5134 "switch_spat_M≔ False " "noBreak"
          global switch_spat_M=  False
        else:
          $ 5136 "ElseIf spatula ≟ 'spatula_S' and switch_spat_S ≟ True and prev_spat≟'spatula_M'" "noBreak"
          if (spatula  ==  "spatula_S" and switch_spat_S  ==   True  and prev_spat == "spatula_M"):
            $ 5137 "MoveL" "noBreak"
            $ 5138 "Spatula_otw" "noBreak"
            movel(Spatula_otw_p, a=1.2, v=0.25)
            $ 5139 "spat_M_up" "noBreak"
            movel(spat_M_up_p, a=1.2, v=0.25)
            $ 5140 "spat_M_pick" "noBreak"
            movel(spat_M_pick_p, a=0.2, v=0.1)
            # begin: URCap Program Node
            #   Source: Robotiq_Grippers, 3.17.0.105337, Robotiq Inc.
            #   Type: Gripper
            $ 5141 "Gripper Open (1)" "noBreak"
            if not(gripper_connected[0]):
              popup("Gripper 1 must be connected to run this program.", "No connection", False, True, True)
            end
            if not(rq_is_gripper_activated("1")):
              popup("Gripper 1 is not activated. Go to Installation tab > Gripper to activate it and run the program again.", "Not activated", False, True, True)
            end
            rq_set_pos_spd_for(0, 255, 77, "1")
            rq_wait_pos_spe_for_request(0, 255, 77, "1")
            rq_go_to("1")
            rq_wait("1")
            # end: URCap Program Node
            $ 5142 "spat_S_pick" "noBreak"
            movel(spat_S_pick_p, a=1.2, v=0.25)
            # begin: URCap Program Node
            #   Source: Robotiq_Grippers, 3.17.0.105337, Robotiq Inc.
            #   Type: Gripper
            $ 5143 "Gripper Close (1)" "noBreak"
            if not(gripper_connected[0]):
              popup("Gripper 1 must be connected to run this program.", "No connection", False, True, True)
            end
            if not(rq_is_gripper_activated("1")):
              popup("Gripper 1 is not activated. Go to Installation tab > Gripper to activate it and run the program again.", "Not activated", False, True, True)
            end
            rq_set_pos_spd_for(255, 0, 77, "1")
            rq_wait_pos_spe_for_request(255, 0, 77, "1")
            rq_go_to("1")
            rq_wait("1")
            # end: URCap Program Node
            $ 5144 "spat_S_up" "noBreak"
            movel(spat_S_up_p, a=1.2, v=0.25)
            $ 5145 "Spatula_otw" "noBreak"
            movel(Spatula_otw_p, a=1.2, v=0.25)
            $ 5146 "switch_spat_S≔ False " "noBreak"
            global switch_spat_S=  False
          else:
            $ 5148 "ElseIf spatula≟'spatula_S' and switch_spat_S≟ True  and prev_spat≟'spatula_L'" "noBreak"
            if (spatula == "spatula_S" and switch_spat_S ==   True    and  prev_spat == "spatula_L"):
              $ 5149 "MoveJ" "noBreak"
              $ 5150 "Spatula_otw" "noBreak"
              movej(get_inverse_kin(Spatula_otw_p, qnear=Spatula_otw_q), a=1.3962634015954636, v=1.0471975511965976)
              $ 5151 "spat_L_up" "noBreak"
              movej(get_inverse_kin(spat_L_up_p, qnear=spat_L_up_q), a=1.3962634015954636, v=1.0471975511965976)
              $ 5152 "MoveL" "noBreak"
              $ 5153 "spat_L_side" "noBreak"
              movel(spat_L_side_p, a=1.2, v=0.25)
              $ 5154 "spat_L_lift" "noBreak"
              movel(spat_L_lift_p, a=1.2, v=0.25)
              $ 5155 "spat_L_pick" "noBreak"
              movel(spat_L_pick_p, a=0.2, v=0.1)
              # begin: URCap Program Node
              #   Source: Robotiq_Grippers, 3.17.0.105337, Robotiq Inc.
              #   Type: Gripper
              $ 5156 "Gripper Open (1)" "noBreak"
              if not(gripper_connected[0]):
                popup("Gripper 1 must be connected to run this program.", "No connection", False, True, True)
              end
              if not(rq_is_gripper_activated("1")):
                popup("Gripper 1 is not activated. Go to Installation tab > Gripper to activate it and run the program again.", "Not activated", False, True, True)
              end
              rq_set_pos_spd_for(0, 255, 77, "1")
              rq_wait_pos_spe_for_request(0, 255, 77, "1")
              rq_go_to("1")
              rq_wait("1")
              # end: URCap Program Node
              $ 5157 "spat_S_pick" "noBreak"
              movel(spat_S_pick_p, a=1.2, v=0.25)
              # begin: URCap Program Node
              #   Source: Robotiq_Grippers, 3.17.0.105337, Robotiq Inc.
              #   Type: Gripper
              $ 5158 "Gripper Close (1)" "noBreak"
              if not(gripper_connected[0]):
                popup("Gripper 1 must be connected to run this program.", "No connection", False, True, True)
              end
              if not(rq_is_gripper_activated("1")):
                popup("Gripper 1 is not activated. Go to Installation tab > Gripper to activate it and run the program again.", "Not activated", False, True, True)
              end
              rq_set_pos_spd_for(255, 0, 77, "1")
              rq_wait_pos_spe_for_request(255, 0, 77, "1")
              rq_go_to("1")
              rq_wait("1")
              # end: URCap Program Node
              $ 5159 "spat_S_up" "noBreak"
              movel(spat_S_up_p, a=1.2, v=0.25)
              $ 5160 "Spatula_otw" "noBreak"
              movel(Spatula_otw_p, a=1.2, v=0.25)
              $ 5161 "switch_spat_S≔ False " "noBreak"
              global switch_spat_S=  False
            else:
              $ 5163 "ElseIf spatula≟'spatula_flat_S'  and switch_spat_F_S ≟ True " "noBreak"
              if (spatula == "spatula_flat_S"   and  switch_spat_F_S  ==   True  ):
                $ 5164 "MoveL" "noBreak"
                $ 5165 "Spatula_otw" "noBreak"
                movel(Spatula_otw_p, a=1.2, v=0.25)
                $ 5166 "spat_flatM_up" "noBreak"
                movel(spat_flatM_up_p, a=1.2, v=0.25)
                $ 5167 "spat_flatM_pick" "noBreak"
                movel(spat_flatM_pick_p, a=0.2, v=0.1)
                # begin: URCap Program Node
                #   Source: Robotiq_Grippers, 3.17.0.105337, Robotiq Inc.
                #   Type: Gripper
                $ 5168 "Gripper Open (1)" "noBreak"
                if not(gripper_connected[0]):
                  popup("Gripper 1 must be connected to run this program.", "No connection", False, True, True)
                end
                if not(rq_is_gripper_activated("1")):
                  popup("Gripper 1 is not activated. Go to Installation tab > Gripper to activate it and run the program again.", "Not activated", False, True, True)
                end
                rq_set_pos_spd_for(0, 255, 74, "1")
                rq_wait_pos_spe_for_request(0, 255, 74, "1")
                rq_go_to("1")
                rq_wait("1")
                # end: URCap Program Node
                $ 5169 "spat_flatS_pick" "noBreak"
                movel(spat_flatS_pick_p, a=1.2, v=0.25)
                # begin: URCap Program Node
                #   Source: Robotiq_Grippers, 3.17.0.105337, Robotiq Inc.
                #   Type: Gripper
                $ 5170 "Gripper Close (1)" "noBreak"
                if not(gripper_connected[0]):
                  popup("Gripper 1 must be connected to run this program.", "No connection", False, True, True)
                end
                if not(rq_is_gripper_activated("1")):
                  popup("Gripper 1 is not activated. Go to Installation tab > Gripper to activate it and run the program again.", "Not activated", False, True, True)
                end
                rq_set_pos_spd_for(255, 0, 77, "1")
                rq_wait_pos_spe_for_request(255, 0, 77, "1")
                rq_go_to("1")
                rq_wait("1")
                # end: URCap Program Node
                $ 5171 "spat_flatS_up" "noBreak"
                movel(spat_flatS_up_p, a=1.2, v=0.25)
                $ 5172 "Spatula_otw" "noBreak"
                movel(Spatula_otw_p, a=1.2, v=0.25)
                $ 5173 "switch_spat_F_S≔ False " "noBreak"
                global switch_spat_F_S=  False
              end
            end
          end
        end
        $ 5175 "Set" "noBreak"
        set_tcp(p[0.0,0.0,0.15052000000000001,3.1415,0.0,0.0])
        $ 5176 "Loop 1 times" "noBreak"
        Loop_9 = 0
        while (Loop_9 < 1):
          $ 5179 "auto_scoop(W_now)" "noBreak"
          auto_scoop(W_now)
          $ 5180 "Wait: 0.5" "noBreak"
          sleep(0.5)
          $ 5181 "Set AO[0]=0.0" "noBreak"
          set_standard_analog_out(0, 0.0)
          Loop_9 = Loop_9 + 1
        end
        $ 5182 "after_scoop_f()" "noBreak"
        after_scoop_f()
        # begin: URCap Program Node
        #   Source: SensoPart VISOR Robotic, 2.0.6, SensoPart Industriesensorik GmbH
        #   Type: Exit Pose
        $ 5183 "Exit Pose" "noBreak"
        movel(pose_trans(easyPickPose,p[0.0000,0.0000,-0.0000,0.0000,0.0000,0.0000]),a=0.5000,v=0.2500,t=0.000000,r=0.000000)
        # end: URCap Program Node
        easyPickObjTaken = True
      end
      # end: URCap Program Node
      # begin: URCap Program Node
      #   Source: SensoPart VISOR Robotic, 2.0.6, SensoPart Industriesensorik GmbH
      #   Type: No Object Detected
      $ 5184 "No Object Detected" "noBreak"
      if (visor_partsFound(easyPickVisorId) < 1):
        $ 5185 "Popup: No weigh scale detected" "noBreak"
        popup("No weigh scale detected", "Message", False, False, blocking=True)
        else:
      end
      # end: URCap Program Node
    end
    easyPickCount_4 = easyPickCount_4 + 1
    visor_easyPickUpdate(easyPickVisorId, "counter", easyPickCount_4)
    visor_easyPickSetIdent("3af2be", easyPickVisorId)
    # end: URCap Program Node
  end
  visorFuncEasyPick_dd8337()
  # end: URCap Program Node
  $ 5186 "Set"
  set_tcp(p[0.0,0.0,0.161,3.1415,0.0,0.0])
